(* IEC 61131-3 sources: Elmo_Master/Lasal_PRG/Elmo_EtherCAT_Test_4Axis/Class/_TCPIPServer, 1 file *)

(* ---- _TCPIPServer.st ---- *)
  #ifndef OS_VERSION_MIN_SALAMANDER
    #define OS_VERSION_MIN_SALAMANDER          0x9000
  #endif
  #define TCP_SVR_NO_ERROR                          0

  #define TCP_SVR_ERR_INVALID_SOCKET            -1

  #define TCP_SVR_ERR_SET_PARA_INVALID_CMD     -10
  #define TCP_SVR_ERR_SET_PARA_INVALID_SUB_CMD -11

  #define TCP_SVR_ERR_TASK_ALREADY_EXIST       -12

  // - RETURN VALUES PRIVATE METHOD Read_AP_TaskPeriod
  #define TCP_SVR_ERR_TASK_TIME_NO_APP            -31
  #define TCP_SVR_ERR_TASK_TIME_WRONG_TASK_TYPE   -33
  #define TCP_SVR_ERR_TASK_TIME_OBJ_NOT_FOUND     -35

  // - RETURN VALUES PRIVATE METHOD Read_LSLOBJ_CRC32
  #define TCP_SVR_ERR_GET_LSLOBJ_NAME             -20
  #define TCP_SVR_ERR_INVALID_POINTER             -21

  // - RETURN VALUES PRIVATE METHOD AP_TaskCreate
  #define TCP_SVR_ERR_TASK_CREATE                 -40

  // - RETURN VALUES PRIVATE METHOD AP_SemaCreate
  #define TCP_SVR_ERR_SEMA_CREATE                 -50
  #define TCP_SVR_ERR_SEMA_INVALID_IDX            -51
  #define TCP_SVR_ERR_SEMA_INVALID_NAME           -52

  #define TCP_SVR_SEND_BUFFER_EMPTY               -6
  #define TCP_SVR_ERR_SEND_BUFFER_FATAL_ERROR     -7

  #define TCP_SVR_SEND_BUFFER_FULL      -4

  #define TCP_SVR_SOCK_INFO_CONNECT                 1
  #define TCP_SVR_SOCK_INFO_DISCONNECT              0

  #define TCP_SVR_ERR_GROUP_OS                      0
  #define TCP_SVR_ERR_GROUP_AP                      1

  #define TCP_SVR_ERR_CODE_AP_TIMEOUT              -1

  #ifndef INIT_FIRSTSCAN
    #define INIT_FIRSTSCAN                         12
  #endif

  #ifndef AP_TASK_PRIORITY_DEFAULT
    #define AP_TASK_PRIORITY_DEFAULT               14
  #endif

  #define TCP_SVR_ERR_MAIN_INIT                   -90

  #define TCP_SVR_ERR_MAX_CONN                    -80

  #ifndef KEEPALIVE_INTERVAL_DEFAULT
    #define KEEPALIVE_INTERVAL_DEFAULT           7200
  #endif

  #ifndef KEEPALIVE_RETRYTIME_DEFAULT
    #define KEEPALIVE_RETRYTIME_DEFAULT            75
  #endif

  #ifndef KEEPALIVE_RETRYCNT_DEFUALT
    #define KEEPALIVE_RETRYCNT_DEFUALT             10
  #endif

  #ifndef CLOSE_SOCKET_TYPE_DEFAULT
    #define CLOSE_SOCKET_TYPE_DEFAULT               0
  #endif

#include "..\..\Class\_TCPIPServer\_TCPIPServer.h"
#include "..\..\Class\_TCPIPServer\SalamanderDelay.h"

(*!
<Class
	Name               = "_TCPIPServer"
	Revision           = "1.2"
	RealtimeTask       = "false"
	CyclicTask         = "true"
	DefCyclictime      = "10 ms"
	BackgroundTask     = "false"
	DefBackground      = "always"
	Sigmatek           = "true"
	OSInterface        = "false"
	HighPriority       = "false"
	Automatic          = "false"
	UpdateMode         = "Prescan"
	SharedCommandTable = "true"
	Objectsize         = "(590,120)"
	Comment            = "TCP/IP Server for TCP/IP Communication">
	<Channels>
		<Server Name="Control" Visualized="false" Initialize="false" WriteProtected="true" Retentive="false" Comment="shows the actual TCP/IP state"/>
		<Server Name="ErrorCode" Visualized="false" Initialize="false" WriteProtected="true" Retentive="false" Comment="Shows error codes&#13;&#10; 0 ... no error&#13;&#10;-1 ... general error&#13;&#10;-2 ... timeout error&#13;&#10;-3 ... connection closed by client&#13;&#10;-4 ... File open failed&#13;&#10;-5 ... Copy Data from File failed&#13;&#10;-6 ... Sending Data failed&#13;&#10;-7 ... read SendBuffer failed&#13;&#10;-8 ... BackUp- or Restore-Object failed&#13;&#10;-9 ... Pointer to SendBuffer = NIL&#13;&#10;-10... Pointer to Receive Buffer = NIL&#13;&#10;-11... Write into SendBuffer failed&#13;&#10;-12... Set Socket Option failed&#13;&#10;-13... Data is to big to send&#13;&#10;-14... Received Data is too short&#13;&#10;-15... Received Datasize not equal with specified Datasize&#13;&#10;-16... Received Datasize not equal with specified Datasize (too long)&#13;&#10;-99... Allocate Memory failed&#13;&#10;-100 . Search for Semikolon or Carriage Return failed"/>
		<Server Name="SemaName01" Visualized="true" Initialize="false" WriteProtected="true" Retentive="false" Comment="name of mutex to save the internal connection buffer&#13;&#10;&#13;&#10;This name is also listed in PLCTraceView"/>
		<Server Name="SemaName02" Visualized="true" Initialize="false" WriteProtected="true" Retentive="false" Comment="name of mutex to save the internal connection settings (socket options)&#13;&#10;&#13;&#10;This name is also listed in PLCTraceView"/>
		<Server Name="TaskName" Visualized="true" Initialize="false" WriteProtected="true" Retentive="false" Comment="shows task information&#13;&#10;-) use object in cyclic task&#13;&#10;-) use object in async task&#13;&#10;-) task deactivated&#13;&#10;-) async task error status (error creating async task)&#13;&#10;&#13;&#10;In case of using the object in async task, this name is also listed in PLCTraceView"/>
		<Client Name="_MultiTask" Required="false" Internal="false" Comment="object channel to OS interface class _MultiTask"/>
		<Client Name="_StdLib" Required="false" Internal="false" Comment="object channel to OS interface class _StdLib"/>
		<Client Name="_TaskObjectControl" Required="false" Internal="false" Comment="object channel to OS interface class _TaskObjectControl"/>
		<Client Name="CheckSum" Required="true" Internal="true"/>
		<Client Name="Config" Required="false" Internal="false" Comment="object configuration&#13;&#10;bit0 ... task configuration&#13;&#10;0 = use object in cyclic task&#13;&#10;1 = use object in async task"/>
		<Client Name="ConnectionsPerRun" Required="true" Internal="false" DefValue="1" Comment="Number of connections to process every cycle:&#13;&#10;&#13;&#10;0, 1 = 1 connection per cycle&#13;&#10;2 = 2 connections per cycle&#13;&#10;... up to ...&#13;&#10;&quot;MaxConnections&quot; = all connections every cycle"/>
		<Client Name="MaxConnections" Required="true" Internal="false" DefValue="0" Comment="Maximal number of connections. Maximal possible connections are 128.&#13;&#10;&#13;&#10;0 = 16 connections, because of compatibility to older versions."/>
		<Client Name="Port" Required="true" Internal="false" Comment="port number&#13;&#10;"/>
		<Client Name="SigCLib" Required="false" Internal="false" Comment="object channel to OS interface class SigCLib"/>
		<Client Name="SizeOfTXBuffer" Required="false" Internal="false" Comment="size of TX buffer [byte]&#13;&#10;if 0 there will be 1024 Byte allocated"/>
		<Client Name="StrSemaName01" Required="true" Internal="true"/>
		<Client Name="StrSemaName02" Required="true" Internal="true"/>
		<Client Name="StrTaskName" Required="true" Internal="true"/>
		<Client Name="Timeout" Required="false" Internal="false" Comment="TCP timeout [ms]&#13;&#10;if 0 then Timeout is deactivated"/>
	</Channels>
	<Dependencies>
		<Files>
			<File Path=".\lsl_st_tcp_user.h" Include="false"/>
			<File Path=".\Class\_TCPIPServer\_TCPIPServer.h" Include="true"/>
			<File Path=".\Class\_TCPIPServer\SalamanderDelay.h" Include="true"/>
		</Files>
	</Dependencies>
	<RevDoku>
		<Owner Company="SIGMATEK"/>
		<Dokumentation Revision="1.2" Date="2024-07-01" Author="zoepat" Company="Sigmatek" Description="- increased maximum connections from 16 to 128.&#13;&#10;- added configuration to define the number of connections to be processed per cycle."/>
		<Dokumentation Revision="1.1" Date="2023-03-23" Author="obechr" Company="Sigmatek" Description="changed comments of parameters for method SendData()"/>
		<Dokumentation Revision="1.0" Date="2019-01-15" Author="hoeant" Company="Sigmatek" Description="creation of class"/>
	</RevDoku>
	<Network Name="_TCPIPServer">
		<!-- List of Components in this network -->
		<Components>
			<Object
				Name       = "CheckSum"
				Class      = "_CheckSum"
				Position   = "(240,180)"
				Visualized = "false">
				<Channels>
					<Server Name="ClassSvr"/>
				</Channels>
			</Object>
			<Object
				Name       = "StrSemaName01"
				Class      = "String"
				Position   = "(240,510)"
				Visualized = "true"
				Remotely   = "true">
				<Channels>
					<Server Name="Data"/>
					<Client Name="SingleRealloc" Value="1"/>
				</Channels>
			</Object>
			<Object
				Name       = "StrSemaName02"
				Class      = "String"
				Position   = "(240,660)"
				Visualized = "true"
				Remotely   = "true">
				<Channels>
					<Server Name="Data"/>
					<Client Name="SingleRealloc" Value="1"/>
				</Channels>
			</Object>
			<Object
				Name       = "StrTaskName"
				Class      = "String"
				Position   = "(240,360)"
				Visualized = "true"
				Remotely   = "true">
				<Channels>
					<Server Name="Data"/>
					<Client Name="SingleRealloc" Value="1"/>
				</Channels>
			</Object>
		</Components>
		<Comments>
		</Comments>
		<!-- List of Connections in this network -->
		<Connections>
			<Connection Source="this.CheckSum" Destination="CheckSum.ClassSvr"/>
			<Connection Source="this.StrTaskName" Destination="StrTaskName.Data"/>
			<Connection Source="this.StrSemaName01" Destination="StrSemaName01.Data"/>
			<Connection Source="this.StrSemaName02" Destination="StrSemaName02.Data"/>
			<Connection Source="this.TaskName" Destination="StrTaskName.Data" Vertices="(1028,330),(556,450),"/>
			<Connection Source="this.SemaName01" Destination="StrSemaName01.Data" Vertices="(1028,390),(556,600),"/>
			<Connection Source="this.SemaName02" Destination="StrSemaName02.Data" Vertices="(1028,450),(556,750),"/>
		</Connections>
		<!-- Headerfiles -->
		<Options>
		</Options>
	</Network>
</Class>
*)
_TCPIPServer : CLASS
	TYPE
#pragma pack(push, 1)
	  _BUFFER : STRUCT  //! <Type Comment="Struct for Receive- and Send-Buffer" Name="_BUFFER"/>
	    udSize : UDINT;  //! <Type Comment="Size of Data" Name="_BUFFER.udSize"/>
	    pData : ^void;  //! <Type Comment="Pointer to Data" Name="_BUFFER.pData"/>
	  END_STRUCT;
#pragma pack(pop)
#pragma pack(push, 1)
	  _BUFFER_HEADER : STRUCT
	    DataSize : UDINT;
	  END_STRUCT;
#pragma pack(pop)
	  _FSM_TCPIP_SERVER :  //! <Type Public="true" Comment="stepping switch for TCP/IP connection" Name="_FSM_TCPIP_SERVER"/>
	  (
	    _STATE_NONE,
	    _STATE_INIT_SERVER,
	    _STATE_NO_USER_INTERFACE_CONNECTED,
	    _STATE_IDLE,
	    _STATE_MAIN_SOCK,
	    _STATE_LISTEN,
	    _STATE_ACCEPT,
	    _STATE_CONNECT,
	    _STATE_RECV,
	    _STATE_SHUTDOWN,
	    _STATE_CLOSE_MAIN_SOCK,
	    _STATE_CLOSE_SOCK,
	    _STATE_ERROR,
	    _STATE_ERROR_ALLOCATING_MEMORY,
	    _STATE_ERROR_CREATING_MUTEX,
	    _STATE_ERROR_CREATING_TASK,
	    _STATE_SEND,
	    _STATE_MAIN_SOCK_OPT,
	    _STATE_DEL_CONNECTION,
	    _STATE_CONN_SOCK_OPT
	  )$UDINT;
#pragma pack(push, 1)
	  _TX_RINGBUFFER : STRUCT  //! <Type Comment="struct to handle a ringbuffer" Name="_TX_RINGBUFFER"/>
	    udSize : UDINT;
	    udUsed : UDINT;
	    pMem : ^void;
	    pRead : ^CHAR;
	    pWrite : ^CHAR;
	  END_STRUCT;
#pragma pack(pop)
	  _SocketOptions : BDINT
	  [
	    1 Nagle,
	    2 KeepAlive,
	    3 DelayedAck,
	    4 ReuseAddr,
	    5 Bit5,
	    6 Bit6,
	    7 Bit7,
	    8 Bit8,
	    9 Bit9,
	    10 Bit10,
	    11 Bit11,
	    12 Bit12,
	    13 Bit13,
	    14 Bit14,
	    15 Bit15,
	    16 Bit16,
	    17 Bit17,
	    18 Bit18,
	    19 Bit19,
	    20 Bit20,
	    21 Bit21,
	    22 Bit22,
	    23 Bit23,
	    24 Bit24,
	    25 Bit25,
	    26 Bit26,
	    27 Bit27,
	    28 Bit28,
	    29 Bit29,
	    30 Bit30,
	    31 Bit31,
	    32 Bit32,
	  ];
#pragma pack(push, 1)
	  _KeepAlivePara : STRUCT
	    keepIDLE : DINT;
	    keepINTVL : DINT;
	    keepCNT : DINT;
	  END_STRUCT;
#pragma pack(pop)
#pragma pack(push, 1)
	  _CONNECTION : STRUCT
	    dSocket : DINT;
	    FSM_TCP : _FSM_TCPIP_SERVER;
	    udTimeStamp : UDINT;
	    SendBuffer : _TX_RINGBUFFER;
	    pBufferWaitForSendig : ^CHAR;
	    pBufferWaitForSendingHelp : ^CHAR;
	    BufferHeader : _BUFFER_HEADER;
	    ConnSockOpt : _SocketOptions;
	    pNextConn : ^_CONNECTION;
	    bdSettings : BDINT
	    [
	      1 SockOptChanged,
	      2 Bit2,
	      3 Bit3,
	      4 Bit4,
	      5 Bit5,
	      6 Bit6,
	      7 Bit7,
	      8 Bit8,
	      9 Bit9,
	      10 Bit10,
	      11 Bit11,
	      12 Bit12,
	      13 Bit13,
	      14 Bit14,
	      15 Bit15,
	      16 Bit16,
	      17 Bit17,
	      18 Bit18,
	      19 Bit19,
	      20 Bit20,
	      21 Bit21,
	      22 Bit22,
	      23 Bit23,
	      24 Bit24,
	      25 Bit25,
	      26 Bit26,
	      27 Bit27,
	      28 Bit28,
	      29 Bit29,
	      30 Bit30,
	      31 Bit31,
	      32 Bit32,
	    ];
	    KeepAlivePara : _KeepAlivePara;
	    CloseSocketType : UDINT;
	  END_STRUCT;
#pragma pack(pop)
#pragma pack(push, 1)
	  _KeepAliveParaLasalOS : STRUCT
	    interval : UINT;
	    retry : UINT;
	    timeout : UINT;
	  END_STRUCT;
#pragma pack(pop)
	END_TYPE
  //Servers:
	Control 	: SvrChCmd__FSM_TCPIP_SERVER_PTofCls__TCPIPServer;
	ErrorCode 	: SvrCh_DINT;
	TaskName 	: SvrCh_UDINT;
	SemaName01 	: SvrCh_UDINT;
	SemaName02 	: SvrCh_UDINT;
  //Clients:
	Port 	: CltCh_DINT;
	Timeout 	: CltCh_DINT;
	SizeOfTXBuffer 	: CltCh_UDINT;
	MaxConnections 	: CltCh_DINT;
	ConnectionsPerRun 	: CltCh_DINT;
	Config 	: CltCh_DINT;
	_StdLib 	: CltChCmd__StdLib;
	_MultiTask 	: CltChCmd__MultiTask;
	SigCLib 	: CltChCmd_SigCLib;
	CheckSum 	: CltChCmd__CheckSum;
	StrTaskName 	: CltChCmd_String;
	StrSemaName01 	: CltChCmd_String;
	StrSemaName02 	: CltChCmd_String;
	_TaskObjectControl 	: CltChCmd__TaskObjectControl;
  //Variables:
		dMainSock 	: DINT;			//! <Variable Comment="main socket for TCP/IP connection" Name="dMainSock"/>
		FSM_TCP 	: _FSM_TCPIP_SERVER;			//! <Variable Comment="finite state machine for TCP/IP connection" Name="FSM_TCP"/>
		SocketArray : ARRAY [0..127] OF _CONNECTION;
			//! <Variable Comment="Saves the Informations for each Connection" Name="SocketArray"/>
		RECVbuffer 	: _BUFFER;			//! <Variable Comment="struct of Receive buffer" Name="RECVbuffer"/>
		lsl_tcp_user 	: ^LSL_TCP_USER;
		usInit 	: USINT;
		bdStatus : BDINT
		[
		  1 SalamanderOS,
		  5 CIL_tcp_user,
		  6 CIL_ssl_user,
		  7 CIL_debug,
		  9 InhibNextConn,
		  13 LSLOBJ_CRC32,
		  14 AP_TaskPeriod,
		  15 CyclicTask,
		  16 AsyncTask,
		  17 Sema01,
		  18 Sema02,
		  25 ErrAsyncTask,
		  26 ErrSema01,
		  27 ErrSema02,
		  28 ErrMem,
		  29 ErrorNoUserInterface,
		];

		MaxConn 	: DINT;
		lsl_ssl_user 	: ^LSL_SSL_USER;
		pCIL_DEBUG 	: ^OS_SALAMANDERDEBUG;
		MainSockOpt 	: _SocketOptions;
		AP_TaskTime 	: UDINT;
		AP_TaskHandle 	: MT_TASKHANDLE;
		AP_SemaHandle1 	: MT_SEMAHANDLE;
		AP_SemaSockOpt 	: MT_SEMAHANDLE;
		ActConn 	: DINT;
		pActConn 	: ^_CONNECTION;
		udTimeStamp 	: UDINT;
		udTimeAccept 	: UDINT;
		AP_TaskPriority 	: UDINT;
		KeepAlivePara 	: _KeepAlivePara;
		CloseSocketType 	: UDINT;
		dNewSock 	: DINT;
		pThisInterface 	: ^_TCPIPServerInterface;
  //Functions:
				//! <Function Comment="-) initialize TCP USER pointer to use OS TCP FUNCTIONS&#13;&#10;-) read port number&#13;&#10;-) Allocate Memory for Buffers" Name="Init"/>
	FUNCTION VIRTUAL GLOBAL Init;
				//! <Function Comment="cyclic tast methode which is called if client &#13;&#10;cConfig = 0" Name="CyWork"/>
	FUNCTION VIRTUAL GLOBAL CyWork
		VAR_INPUT
			EAX 	: UDINT;
		END_VAR
		VAR_OUTPUT
			state (EAX) 	: UDINT;
		END_VAR;
				//! <Function Comment="this function writes data into the TX buffer&#13;&#10;" Name="SENDbuffer_Write"/>
	FUNCTION SENDbuffer_Write
		VAR_INPUT
			pData 	: ^void;
			udSize 	: UDINT;
			pBuffer 	: ^_TX_RINGBUFFER;
		END_VAR
		VAR_OUTPUT
			dRetcode 	: DINT;
		END_VAR;
				//! <Function Comment="Function to send data over TCP/IP&#13;&#10;&#13;&#10;--------------------------------------&#13;&#10;Input variables&#13;&#10;--------------------------------------&#13;&#10;-) pData ... pointer to data to send&#13;&#10;-) udSize ... size of data to send [byte]&#13;&#10;-) dSock ... Receiver-Socket&#13;&#10;&#13;&#10;--------------------------------------&#13;&#10;Output variables&#13;&#10;--------------------------------------&#13;&#10;-) dRetcode&#13;&#10;   &lt; 0:&#13;&#10;      -1 ... TCP Client not ready&#13;&#10;      else ... OS TCP error code&#13;&#10;&#13;&#10;   &gt;=0:&#13;&#10;      dRetcode = udSize ... Sending data over TCP/IP successful" Name="SendTCP"/>
	FUNCTION SendTCP
		VAR_INPUT
			pData 	: ^void;
			udSize 	: UDINT;
			dSock 	: DINT;
			bDirect 	: DINT;
		END_VAR
		VAR_OUTPUT
			dRetcode 	: DINT;
		END_VAR;
				//! <Function Comment="Handles the Connection and Data receiving and sending" Name="CyclicCall"/>
	FUNCTION VIRTUAL GLOBAL CyclicCall;
				//! <Function Comment="Read Send Buffer" Name="SENDbuffer_Read"/>
	FUNCTION SENDbuffer_Read
		VAR_INPUT
			pBuffer 	: ^_TX_RINGBUFFER;
			pData 	: ^void;
			udSize 	: UDINT;
		END_VAR
		VAR_OUTPUT
			Retcode 	: DINT;
		END_VAR;
				//! <Function Comment="Send Data over TCP/IP" Name="SendData"/>
	FUNCTION VIRTUAL GLOBAL SendData
		VAR_INPUT
			pData 	: ^void;			//! <Variable Comment="Pointer to Data" Name="SendData.pData"/>
			udSize 	: UDINT;			//! <Variable Comment="Size of Data" Name="SendData.udSize"/>
			dSock 	: DINT;			//! <Variable Comment="Socket to which it should be send" Name="SendData.dSock"/>
			bDirect 	: BOOL;			//! <Variable Comment="0 ... Write it to Send Buffer and send it in next Cyclus&#13;&#10;1 ... Send it imediatly" Name="SendData.bDirect"/>
		END_VAR
		VAR_OUTPUT
			dRetcode 	: DINT;			//! <Variable Comment="&gt;=0 .. size of the processed data&#13;&#10;&lt;0 ..  error occured" Name="SendData.dRetcode"/>
		END_VAR;

	FUNCTION Read_LSLOBJ_CRC32
		VAR_INPUT
			pCRC32 	: ^CHAR;
		END_VAR
		VAR_OUTPUT
			Retcode 	: DINT;
		END_VAR;

	FUNCTION Read_AP_TaskPeriod
		VAR_OUTPUT
			Retcode 	: DINT;
		END_VAR;

	FUNCTION AP_TaskCreate
		VAR_INPUT
			pTaskName 	: ^CHAR;
			pCallback 	: ^void;
		END_VAR
		VAR_OUTPUT
			Retcode 	: DINT;
		END_VAR;

	FUNCTION AP_TaskCallback
		VAR_INPUT
			Param0 	: ^void;
		END_VAR;

	FUNCTION GetMultiTaskErrorCode
		VAR_INPUT
			pErrTxt 	: ^CHAR;
		END_VAR;

	FUNCTION AP_SemaCreate
		VAR_INPUT
			pSemaName 	: ^CHAR;
			Index 	: DINT;
		END_VAR
		VAR_OUTPUT
			Retcode 	: DINT;
		END_VAR;

	FUNCTION AP_TaskDelay
		VAR_INPUT
			udTaskDelay 	: UDINT;
		END_VAR;

	FUNCTION SetMainSocketOptions
		VAR_OUTPUT
			Retcode 	: DINT;
		END_VAR;

	FUNCTION RingbufferReadEntry
		VAR_INPUT
			pBuffer 	: ^_TX_RINGBUFFER;
			pData 	: ^void;
			pSize 	: ^UDINT;
		END_VAR
		VAR_OUTPUT
			Retcode 	: DINT;
		END_VAR;

	FUNCTION RingbufferWriteEntry
		VAR_INPUT
			pBuffer 	: ^_TX_RINGBUFFER;
			pData 	: ^void;
			udSize 	: UDINT;
		END_VAR
		VAR_OUTPUT
			Retcode 	: DINT;
		END_VAR;

	FUNCTION AP_SemaWait
		VAR_INPUT
			SemaHandle 	: MT_SEMAHANDLE;
		END_VAR;

	FUNCTION AP_SemaSignal
		VAR_INPUT
			SemaHandle 	: MT_SEMAHANDLE;
		END_VAR;

	FUNCTION SetSocketOptions
		VAR_INPUT
			pConn 	: ^_CONNECTION;
		END_VAR
		VAR_OUTPUT
			Retcode 	: DINT;
		END_VAR;

	FUNCTION AddConnIntern
		VAR_INPUT
			dSocket 	: DINT;
			ppConn 	: ^pVoid;
		END_VAR
		VAR_OUTPUT
			Retcode 	: DINT;
		END_VAR;

	FUNCTION DelConnIntern
		VAR_INPUT
			dSocket 	: DINT;
		END_VAR
		VAR_OUTPUT
			Retcode 	: DINT;
		END_VAR;
				//! <Function Comment="method is called with socket informations of the connection sockets" Name="ConnSocketInfo"/>
	FUNCTION ConnSocketInfo
		VAR_INPUT
			dSock 	: DINT;			//! <Variable Comment="socket number" Name="ConnSocketInfo.dSock"/>
			InfoPara1 	: DINT;			//! <Variable Comment="0 ... socket disconnected&#13;&#10;1 ... socket connected" Name="ConnSocketInfo.InfoPara1"/>
			InfoPara2 	: DINT;			//! <Variable Comment="InfoPara2 = 0" Name="ConnSocketInfo.InfoPara2"/>
		END_VAR;
				//! <Function Comment="method is called with socket error status of the connection sockets&#13;&#10;&#13;&#10;-) TCP error (callback: ErrorGroup = 0, ErrorCode = TCP error status)&#13;&#10;-) error code definition in lsl_st_tcp_user.h&#13;&#10;&#13;&#10;-)  internal error (callback: ErrorGroup = 1, ErrorCode = internal error status)&#13;&#10;-) -1: receive timeout (in case of timeout is set)" Name="ConnSocketError"/>
	FUNCTION ConnSocketError
		VAR_INPUT
			dSock 	: DINT;			//! <Variable Comment="socket number" Name="ConnSocketError.dSock"/>
			FSM_TCP 	: _FSM_TCPIP_SERVER;			//! <Variable Comment="status of the state machine of the connection socket" Name="ConnSocketError.FSM_TCP"/>
			ErrGroup 	: DINT;			//! <Variable Comment="0 ... OS error (OS_TCP_USER)&#13;&#10;1 ... AP error (connection timeout)" Name="ConnSocketError.ErrGroup"/>
			ErrCode 	: DINT;			//! <Variable Comment="ErrGroup = 0 (OS error)&#13;&#10;ErrCode definition in lsl_st_tcp_user.h&#13;&#10;&#13;&#10;ErrGroup = 1 (AP error)&#13;&#10;ErrCode = -1 ... connection timeout&#13;&#10;" Name="ConnSocketError.ErrCode"/>
		END_VAR;
				//! <Function Comment="method is called with socket informations of the main socket" Name="MainSocketError"/>
	FUNCTION MainSocketError
		VAR_INPUT
			FSM_TCP 	: _FSM_TCPIP_SERVER;			//! <Variable Comment="status of the state machine of the main socket" Name="MainSocketError.FSM_TCP"/>
			ErrGroup 	: DINT;			//! <Variable Comment="0 ... OS error (OS_TCP_USER)" Name="MainSocketError.ErrGroup"/>
			ErrCode 	: DINT;
		END_VAR;
				//! <Function Comment="Method to set main parameters. Main parameters will be used for every new connection." Name="SetMainParameter"/>
	FUNCTION VIRTUAL GLOBAL SetMainParameter
		VAR_INPUT
			Cmd 	: DINT;			//! <Variable Comment="0 ... (SVR_TCP_CMD_SETSOCKOPT) socket option&#13;&#10;1 ... (SVR_TCP_CMD_TASKPRIO) task priority of async task (in case of using object in async task)&#13;&#10;2 ... (SVR_TCP_CMD_CLOSESOCKETTYPE) close socket type&#13;&#10;3 ... (SVR_TCP_CMD_KEEPALIVEPARA) keep alive parameter&#13;&#10;" Name="SetMainParameter.Cmd"/>
			SubCmd 	: DINT;			//! <Variable Comment="Cmd = 0 (SVR_TCP_CMD_SETSOCKOPT)&#13;&#10;-) SubCmd = 0:  SVR_TCP_SOCKOPT_NAGLE ... activate/deactivate nagle algorithm&#13;&#10;-) SubCmd = 1:  SVR_TCP_SOCKOPT_KEEPALIVE ... activate/deactivate keepalive message&#13;&#10;-) SubCmd = 2:  SVR_TCP_SOCKOPT_DELAYEDACK ... activate/deactivate delayed acknowledge packet&#13;&#10;-) SubCmd = 3:  SVR_TCP_SOCKOPT_REUSEADDR ... activate/deactivate option reuse address&#13;&#10;&#13;&#10;Cmd = 1 (SVR_TCP_CMD_TASKPRIO)&#13;&#10;-) SubCmd = 0: task priority of async task&#13;&#10;&#13;&#10;&#13;&#10;Cmd = 2 (SVR_TCP_CMD_CLOSESOCKETTYPE)&#13;&#10;-) SubCmd = 0: SVR_TCP_CLOSESOCKETTYPE&#13;&#10;&#13;&#10;Cmd = 3 (SVR_TCP_CMD_KEEPALIVEPARA)&#13;&#10;-) SubCmd = 0:  SVR_TCP_KEEPALIVE_KEEPIDLE&#13;&#10;-) SubCmd = 1:  SVR_TCP_KEEPALIVE_KEEPINTVL&#13;&#10;-) SubCmd = 2:  SVR_TCP_KEEPALIVE_KEEPCNT&#13;&#10;" Name="SetMainParameter.SubCmd"/>
			ParaValue 	: DINT;			//! <Variable Comment="Cmd = 0 (SVR_TCP_CMD_SETSOCKOPT)&#13;&#10;-) 1 ... Activate option&#13;&#10;-) 0 ... Deactivate option&#13;&#10;&#13;&#10;Cmd = 1 (SVR_TCP_CMD_TASKPRIO)&#13;&#10;-) task priority 1-14&#13;&#10;&#13;&#10;Cmd = 2 (SVR_TCP_CMD_CLOSESOCKETTYPE)&#13;&#10;-) 0 ... Graceful Close&#13;&#10;-) 1 ... Hard Close&#13;&#10;&#13;&#10;Cmd = 3 (SVR_TCP_CMD_KEEPALIVEPARA)&#13;&#10;-)SubCmd = 0: Interval time [ms] for the Keep Alive packages&#13;&#10;-)SubCmd = 1: Retry time [ms] of Keep Alive packages&#13;&#10;-)SubCmd = 2: Define how often the retry will be attempted. Retry time * Retry Count = timeout for Keep Alive packages" Name="SetMainParameter.ParaValue"/>
		END_VAR
		VAR_OUTPUT
			Retcode 	: DINT;			//! <Variable Comment="0 ... success&#13;&#10;-10 ... invalid CMD&#13;&#10;-11 ... invalid SubCMD&#13;&#10;-12 ... error set task priority - task already created&#13;&#10;-90 ... object not initialized (initialization in first Init() call)" Name="SetMainParameter.Retcode"/>
		END_VAR;
				//! <Function Comment="method to read main parameters" Name="ReadMainParameter"/>
	FUNCTION VIRTUAL GLOBAL ReadMainParameter
		VAR_INPUT
			Cmd 	: DINT;			//! <Variable Comment="0 ... (SVR_TCP_CMD_SETSOCKOPT) socket option&#13;&#10;1 ... (SVR_TCP_CMD_TASKPRIO) task priority of async task (in case of using object in async task)&#13;&#10;2 ... (SVR_TCP_CMD_CLOSESOCKETTYPE) close socket type&#13;&#10;3 ... (SVR_TCP_CMD_KEEPALIVEPARA) keep alive parameter" Name="ReadMainParameter.Cmd"/>
			SubCmd 	: DINT;			//! <Variable Comment="Cmd = 0 (SVR_TCP_CMD_SETSOCKOPT)&#13;&#10;-) SubCmd = 0:  SVR_TCP_SOCKOPT_NAGLE ... activate/deactivate nagle algorithm&#13;&#10;-) SubCmd = 1:  SVR_TCP_SOCKOPT_KEEPALIVE ... activate/deactivate keepalive message&#13;&#10;-) SubCmd = 2:  SVR_TCP_SOCKOPT_DELAYEDACK ... activate/deactivate delayed acknowledge packet&#13;&#10;-) SubCmd = 3:  SVR_TCP_SOCKOPT_REUSEADDR ... activate/deactivate option reuse address&#13;&#10;&#13;&#10;Cmd = 1 (SVR_TCP_CMD_TASKPRIO)&#13;&#10;-) SubCmd = 0: task priority of async task&#13;&#10;&#13;&#10;&#13;&#10;Cmd = 2 (SVR_TCP_CMD_CLOSESOCKETTYPE)&#13;&#10;-) SubCmd = 0: SVR_TCP_CLOSESOCKETTYPE&#13;&#10;&#13;&#10;Cmd = 3 (SVR_TCP_CMD_KEEPALIVEPARA)&#13;&#10;-) SubCmd = 0:  SVR_TCP_KEEPALIVE_KEEPIDLE&#13;&#10;-) SubCmd = 1:  SVR_TCP_KEEPALIVE_KEEPINTVL&#13;&#10;-) SubCmd = 2:  SVR_TCP_KEEPALIVE_KEEPCNT&#13;&#10;" Name="ReadMainParameter.SubCmd"/>
			pParaValue 	: ^DINT;			//! <Variable Comment="pointer to target parameter value" Name="ReadMainParameter.pParaValue"/>
		END_VAR
		VAR_OUTPUT
			Retcode 	: DINT;			//! <Variable Comment="0 ... success&#13;&#10;-10 ... invalid CMD&#13;&#10;-11 ... invalid SubCMD&#13;&#10;-90 ... object not initialized (initialization in first Init() call)" Name="ReadMainParameter.Retcode"/>
		END_VAR;
				//! <Function Comment="method to set connection socket parameters" Name="SetSocketParameter"/>
	FUNCTION VIRTUAL GLOBAL SetSocketParameter
		VAR_INPUT
			dSock 	: DINT;			//! <Variable Comment="socket number" Name="SetSocketParameter.dSock"/>
			Cmd 	: DINT;			//! <Variable Comment="0 ... (SVR_TCP_CMD_SETSOCKOPT) socket option&#13;&#10;2 ... (SVR_TCP_CMD_CLOSESOCKETTYPE) close socket type&#13;&#10;3 ... (SVR_TCP_CMD_KEEPALIVEPARA) keep alive parameter" Name="SetSocketParameter.Cmd"/>
			SubCmd 	: DINT;			//! <Variable Comment="Cmd = 0 (SVR_TCP_CMD_SETSOCKOPT)&#13;&#10;-) SubCmd = 0:  SVR_TCP_SOCKOPT_NAGLE ... activate/deactivate nagle algorithm&#13;&#10;-) SubCmd = 1:  SVR_TCP_SOCKOPT_KEEPALIVE ... activate/deactivate keepalive message&#13;&#10;-) SubCmd = 2:  SVR_TCP_SOCKOPT_DELAYEDACK ... activate/deactivate delayed acknowledge packet&#13;&#10;-) SubCmd = 3:  SVR_TCP_SOCKOPT_REUSEADDR ... activate/deactivate option reuse address&#13;&#10;&#13;&#10;Cmd = 2 (SVR_TCP_CMD_CLOSESOCKETTYPE)&#13;&#10;-) SubCmd = 0: SVR_TCP_CLOSESOCKETTYPE&#13;&#10;&#13;&#10;Cmd = 3 (SVR_TCP_CMD_KEEPALIVEPARA)&#13;&#10;-) SubCmd = 0:  SVR_TCP_KEEPALIVE_KEEPIDLE&#13;&#10;-) SubCmd = 1:  SVR_TCP_KEEPALIVE_KEEPINTVL&#13;&#10;-) SubCmd = 2:  SVR_TCP_KEEPALIVE_KEEPCNT&#13;&#10;" Name="SetSocketParameter.SubCmd"/>
			ParaValue 	: DINT;			//! <Variable Comment="Cmd = 0 (socket option)&#13;&#10;-) 1 ... Activate option&#13;&#10;-) 0 ... Deactivate option&#13;&#10;&#13;&#10;Cmd = 2 (SVR_TCP_CMD_CLOSESOCKETTYPE)&#13;&#10;-) 0 ... Graceful Close&#13;&#10;-) 1 ... Hard Close&#13;&#10;&#13;&#10;Cmd = 3 (SVR_TCP_CMD_KEEPALIVEPARA)&#13;&#10;-)SubCmd = 0: Interval time [ms] for the Keep Alive packages&#13;&#10;-)SubCmd = 1: Retry time [ms] of Keep Alive packages&#13;&#10;-)SubCmd = 2: Define how often the retry will be attempted. Retry time * Retry Count = timeout for Keep Alive packages" Name="SetSocketParameter.ParaValue"/>
		END_VAR
		VAR_OUTPUT
			Retcode 	: DINT;			//! <Variable Comment="0 ... success&#13;&#10;-1 ... invalid socket number&#13;&#10;-10 ... invalid CMD&#13;&#10;-11 ... invalid SubCMD" Name="SetSocketParameter.Retcode"/>
		END_VAR;
				//! <Function Comment="method to read connection socket parameters" Name="ReadSocketParameter"/>
	FUNCTION VIRTUAL GLOBAL ReadSocketParameter
		VAR_INPUT
			dSock 	: DINT;			//! <Variable Comment="socket number" Name="ReadSocketParameter.dSock"/>
			Cmd 	: DINT;			//! <Variable Comment="0 ... (SVR_TCP_CMD_SETSOCKOPT) socket option&#13;&#10;2 ... (SVR_TCP_CMD_CLOSESOCKETTYPE) close socket type&#13;&#10;3 ... (SVR_TCP_CMD_KEEPALIVEPARA) keep alive parameter" Name="ReadSocketParameter.Cmd"/>
			SubCmd 	: DINT;			//! <Variable Comment="Cmd = 0 (SVR_TCP_CMD_SETSOCKOPT)&#13;&#10;-) SubCmd = 0:  SVR_TCP_SOCKOPT_NAGLE ... activate/deactivate nagle algorithm&#13;&#10;-) SubCmd = 1:  SVR_TCP_SOCKOPT_KEEPALIVE ... activate/deactivate keepalive message&#13;&#10;-) SubCmd = 2:  SVR_TCP_SOCKOPT_DELAYEDACK ... activate/deactivate delayed acknowledge packet&#13;&#10;-) SubCmd = 3:  SVR_TCP_SOCKOPT_REUSEADDR ... activate/deactivate option reuse address&#13;&#10;&#13;&#10;Cmd = 2 (SVR_TCP_CMD_CLOSESOCKETTYPE)&#13;&#10;-) SubCmd = 0: SVR_TCP_CLOSESOCKETTYPE&#13;&#10;&#13;&#10;Cmd = 3 (SVR_TCP_CMD_KEEPALIVEPARA)&#13;&#10;-) SubCmd = 0:  SVR_TCP_KEEPALIVE_KEEPIDLE&#13;&#10;-) SubCmd = 1:  SVR_TCP_KEEPALIVE_KEEPINTVL&#13;&#10;-) SubCmd = 2:  SVR_TCP_KEEPALIVE_KEEPCNT&#13;&#10;" Name="ReadSocketParameter.SubCmd"/>
			pParaValue 	: ^DINT;			//! <Variable Comment="pointer to target parameter value" Name="ReadSocketParameter.pParaValue"/>
		END_VAR
		VAR_OUTPUT
			Retcode 	: DINT;			//! <Variable Comment="0 ... success&#13;&#10;-1 ... invalid socket number&#13;&#10;-10 ... invalid CMD&#13;&#10;-11 ... invalid SubCMD" Name="ReadSocketParameter.Retcode"/>
		END_VAR;

	FUNCTION CheckSocketValid
		VAR_INPUT
			dSock 	: DINT;
			ppConn 	: ^pVoid;
		END_VAR
		VAR_OUTPUT
			Retcode 	: BOOL;
		END_VAR;
				//! <Function Comment="Internal Methode to register the Interface Object." Name="AddInterface"/>
	FUNCTION GLOBAL AddInterface
		VAR_INPUT
			thispointer 	: ^void;			//! <Variable Comment="pointer to InterfaceObjekt (this)&#13;&#10;" Name="AddInterface.thispointer"/>
		END_VAR
		VAR_OUTPUT
			dRetcode 	: DINT;			//! <Variable Comment="1..OK (Interface installed )&#13;&#10;-1.. Error (Interface already installed)&#13;&#10;-2.. Error (Pointer not valid)" Name="AddInterface.dRetcode"/>
		END_VAR;
  //Tables:
	FUNCTION @STD
		VAR_OUTPUT
			ret_code	: CONFSTATES;
		END_VAR;
	FUNCTION GLOBAL TAB @CT_;
END_CLASS;

#pragma using _CheckSum
#pragma using String
#pragma usingLtd _MultiTask
#pragma usingLtd _StdLib
#pragma usingLtd _TaskObjectControl
#pragma usingLtd SigCLib

#pragma usingLtd _TCPIPServerInterface

#pragma usingltd _TCPIPServerInterface

FUNCTION VIRTUAL GLOBAL _TCPIPServer::Init
VAR
	i                     : USINT;
  udStrLen              : UDINT;
  dRet                  : DINT;
  szCRC32               : ARRAY [0..15] OF CHAR;
  szTaskName            : ARRAY [0..63] OF CHAR;
  szErrCode             : ARRAY [0..31] OF CHAR;
  szSemaName            : ARRAY [0..63] OF CHAR;
END_VAR

  // -------------------------------------------------------------------------------------------------------
  // -------------------------------------------------------------------------------------------------------
  // - F I R S T   I N I T   R U N   ( M A I N   I N I T )
  // -------------------------------------------------------------------------------------------------------
  // -------------------------------------------------------------------------------------------------------
  FSM_TCP := _STATE_INIT_SERVER;
  if (usInit = 0) then

    // -------------------------------------------------------------------------------------
    // -------------------------------------------------------------------------------------
    // - SET DEFAULT SETTINGS
    // -------------------------------------------------------------------------------------
    // -------------------------------------------------------------------------------------
    MainSockOpt.Nagle      := true;
    MainSockOpt.KeepAlive  := false;
    MainSockOpt.DelayedAck := true;
    MainSockOpt.ReuseAddr  := true;

    AP_TaskPriority         := AP_TASK_PRIORITY_DEFAULT;

    KeepAlivePara.keepIDLE  := KEEPALIVE_INTERVAL_DEFAULT;
    KeepAlivePara.keepINTVL := KEEPALIVE_RETRYTIME_DEFAULT;
    KeepAlivePara.keepCNT   := KEEPALIVE_RETRYCNT_DEFUALT;

    CloseSocketType         := CLOSE_SOCKET_TYPE_DEFAULT;

    // -------------------------------------------------------------------------------------
    // -------------------------------------------------------------------------------------
    // - READ CONFIGURATION PARAMETER
    // -------------------------------------------------------------------------------------
    // -------------------------------------------------------------------------------------
    Port           := Port.Read();
    Config         := Config.Read();
    Timeout        := Timeout.Read();
    MaxConnections := MaxConnections.Read();
    SizeOfTXBuffer := SizeOfTXBuffer.Read();
    ConnectionsPerRun := ConnectionsPerRun.Read();

    // -------------------------------------------------------------------------------------
    // -------------------------------------------------------------------------------------
    // - CHECK GENERAL PARAMETER CONFIGURATION
    // -------------------------------------------------------------------------------------
    // -------------------------------------------------------------------------------------
    if MaxConnections <= 0 then
      MaxConnections := 16;
    elsif MaxConnections > 128 then
      MaxConnections := 128;
    end_if;
    MaxConn := MaxConnections;

    if (SizeOfTXBuffer = 0) then
      SizeOfTXBuffer := 1024;
    end_if;

    //limit between 1 and MaxConnections
    if ConnectionsPerRun <= 0 then
      ConnectionsPerRun := 1;
    elsif ConnectionsPerRun > MaxConnections then
      ConnectionsPerRun := MaxConnections;
    end_if;

    // -------------------------------------------------------------------------------------
    // -------------------------------------------------------------------------------------
    // - READ OS INFORMATION
    // -------------------------------------------------------------------------------------
    // -------------------------------------------------------------------------------------
    if (_RtOSVersion >= OS_VERSION_MIN_SALAMANDER) then
      bdStatus.SalamanderOS := true;
    end_if;

    // -------------------------------------------------------------------------------------
    // -------------------------------------------------------------------------------------
    // - READ OS CIL INTERFACE INFORMATION
    // -------------------------------------------------------------------------------------
    // -------------------------------------------------------------------------------------
    if OS_CILGET("TCP_USER", #lsl_tcp_user) then
      lsl_tcp_user := NIL;
    else
      bdStatus.CIL_tcp_user := true;
    end_if;

    if OS_CILGET("SSL_USER", #lsl_ssl_user) then
      lsl_ssl_user := NIL;
    else
      bdStatus.CIL_ssl_user := true;
    end_if;

    if OS_CILGET("SALAMANDERDEBUG", #pCIL_DEBUG) then
      pCIL_DEBUG := NIL;
    else
      bdStatus.CIL_debug := true;
    end_if;

    // -------------------------------------------------------------------------------------
    // -------------------------------------------------------------------------------------
    // - ALLOCATE MEMORY FOR RECEIVE BUFFER
    // -------------------------------------------------------------------------------------
    // -------------------------------------------------------------------------------------
    RECVbuffer.pData := _StdLib.Malloc(size := to_UDINT(SizeOfTXBuffer));
    if (RECVbuffer.pData = NIL) then
      bdStatus.ErrMem := true;
      ErrorCode := -99;
    end_if;

    // -------------------------------------------------------------------------------------
    // -------------------------------------------------------------------------------------
    // - ALLOCATE MEMORY FOR SEND BUFFER
    // -------------------------------------------------------------------------------------
    // -------------------------------------------------------------------------------------
    for i := 0 to ((MaxConn-1)$USINT) do

      SocketArray[i].dSocket     := 0;
      SocketArray[i].udTimeStamp := 0;
      SocketArray[i].FSM_TCP     := _STATE_IDLE;
      SocketArray[i].pNextConn   := NIL;
      SocketArray[i].SendBuffer.pMem := _StdLib.Malloc(size:=(SizeOfTXBuffer + (10 *sizeof(_BUFFER_HEADER)))); // allocate memory for Ringbuffer (+ 10 * size of Buffer-Header to have enogh Memory)

      if SocketArray[i].SendBuffer.pMem = NIL then
        bdStatus.ErrMem := true;
        ErrorCode := -99;
      else
        SocketArray[i].SendBuffer.pRead  := SocketArray[i].SendBuffer.pMem$^USINT;
        SocketArray[i].SendBuffer.pWrite := SocketArray[i].SendBuffer.pMem$^USINT;
        SocketArray[i].SendBuffer.udSize := SizeOfTXBuffer;
        SocketArray[i].SendBuffer.udUsed := 0;
      end_if;

      SocketArray[i].pBufferWaitForSendig$^void := _StdLib.Malloc(size:=SizeOfTXBuffer); //allocate memory for Sendbuffer

      if SocketArray[i].pBufferWaitForSendig = NIL then
        bdStatus.ErrMem := true;
        ErrorCode := -99;
      end_if;

    end_for;

    // -------------------------------------------------------------------------------------
    // -------------------------------------------------------------------------------------
    // - CHECK USER INTERFACE AVAILABLE
    // -------------------------------------------------------------------------------------
    // -------------------------------------------------------------------------------------

    bdStatus.ErrorNoUserInterface := TRUE;

  end_if;

  usInit += 1;

  // -------------------------------------------------------------------------------------------------------
  // -------------------------------------------------------------------------------------------------------
  // - F I R S T S C A N
  // -------------------------------------------------------------------------------------------------------
  // -------------------------------------------------------------------------------------------------------
  if (_firstscan) then

    // -------------------------------------------------------------------------------------
    // -------------------------------------------------------------------------------------
    // - READ THE LASAL OBJECT CRC32
    // -------------------------------------------------------------------------------------
    // -------------------------------------------------------------------------------------
    dRet := Read_LSLOBJ_CRC32(#szCRC32[0]);
    case dRet of
      (*==================================================================*)
      TCP_SVR_NO_ERROR: // - NO ERROR
      (*==================================================================*)
        bdStatus.LSLOBJ_CRC32 := true;
      (*==================================================================*)
      else // - ERROR WHILE READING THE LASAL OBJECT CRC32 (USE THIS PTR)
      (*==================================================================*)
        SigCLib.IToA(this$DINT, #szCRC32[0], 0x10);
    end_case;

    // -------------------------------------------------------------------------------------
    // -------------------------------------------------------------------------------------
    // - MUTEX CONNECTION INIT
    // -------------------------------------------------------------------------------------
    // -------------------------------------------------------------------------------------
    SigCLib.StrCpy(#szSemaName[0], "USR_SEMA_");
    SigCLib.StrCat(#szSemaName[0], #szCRC32[0]);
    SigCLib.StrCat(#szSemaName[0], "_01");
    dRet := AP_SemaCreate(#szSemaName[4], 0);
    if (dRet = TCP_SVR_NO_ERROR) then
      bdStatus.Sema01 := true;
    else
      bdStatus.ErrSema01 := true;
      GetMultiTaskErrorCode(#szErrCode[0]);
      SigCLib.StrCpy(#szTaskName[0], "SEMA ERR: CREATE SEMA (");
      SigCLib.StrCat(#szTaskName[0], #szErrCode[0]);
      SigCLib.StrCat(#szTaskName[0], ")");
    end_if;

    udStrLen := SigCLib.StrLen(#szSemaName[0]);
    StrSemaName01.WriteDataOff(udStrLen, 0, #szSemaName[0]);

    // -------------------------------------------------------------------------------------
    // -------------------------------------------------------------------------------------
    // - MUTEX SOCKET OPTION INIT
    // -------------------------------------------------------------------------------------
    // -------------------------------------------------------------------------------------
    SigCLib.StrCpy(#szSemaName[0], "USR_SEMA_");
    SigCLib.StrCat(#szSemaName[0], #szCRC32[0]);
    SigCLib.StrCat(#szSemaName[0], "_02");
    dRet := AP_SemaCreate(#szSemaName[4], 1);
    if (dRet = TCP_SVR_NO_ERROR) then
      bdStatus.Sema01 := true;
    else
      bdStatus.ErrSema01 := true;
      GetMultiTaskErrorCode(#szErrCode[0]);
      SigCLib.StrCpy(#szTaskName[0], "SEMA ERR: CREATE SEMA (");
      SigCLib.StrCat(#szTaskName[0], #szErrCode[0]);
      SigCLib.StrCat(#szTaskName[0], ")");
    end_if;

    udStrLen := SigCLib.StrLen(#szSemaName[0]);
    StrSemaName02.WriteDataOff(udStrLen, 0, #szSemaName[0]);

    // -------------------------------------------------------------------------------------
    // -------------------------------------------------------------------------------------
    // - TASK INIT
    // -------------------------------------------------------------------------------------
    // -------------------------------------------------------------------------------------
    udTimeAccept := 500;

    dRet := Read_AP_TaskPeriod();
    if (dRet = TCP_SVR_NO_ERROR) then
      bdStatus.AP_TaskPeriod := true;
      if (Config AND 0x1) then
        // - CYCLIC CALL IN PARALLEL TASK
        SigCLib.StrCpy(#szTaskName[0], "USR_TASK_");
        SigCLib.StrCat(#szTaskName[0], #szCRC32[0]);
        dRet := AP_TaskCreate(#szTaskName[4], #AP_TaskCallback());
        if (dRet = TCP_SVR_NO_ERROR) then
          bdStatus.AsyncTask := true;
        else
          bdStatus.ErrAsyncTask := true;
          GetMultiTaskErrorCode(#szErrCode[0]);
          SigCLib.StrCpy(#szTaskName[0], "TASK ERR: CREATE TASK (");
          SigCLib.StrCat(#szTaskName[0], #szErrCode[0]);
          SigCLib.StrCat(#szTaskName[0], ")");
        end_if;
      else
        // - CYCLIC CALL IN CYCLIC TASK
        bdStatus.CyclicTask := true;
        SigCLib.StrCpy(#szTaskName[0], "CyclicTask");
      end_if;

      // ---------------------------------------------------------------------
      // - ADJUST TIME BETWEEN ACCEPT STEPS FOR COMPATIBILITY
      // ---------------------------------------------------------------------
      if (bdStatus.SalamanderOS = true) then
        udTimeAccept := AP_TaskTime / 1000;
        if (udTimeAccept = 0) then
          udTimeAccept := 1;
        end_if;
      else
        udTimeAccept := AP_TaskTime;
      end_if;
      udTimeAccept := udTimeAccept * 4;

    else

      case dRet of
        (*==================================================================*)
        TCP_SVR_ERR_TASK_TIME_NO_APP:
        (*==================================================================*)
          SigCLib.StrCpy(#szTaskName[0], "TASK ERR: LSLOBJ (NO APPLICATION)");
        (*==================================================================*)
        TCP_SVR_ERR_TASK_TIME_WRONG_TASK_TYPE:
        (*==================================================================*)
          SigCLib.StrCpy(#szTaskName[0], "TASK ERR: LSLOBJ (WRONG TASK TYPE)");
        (*==================================================================*)
        TCP_SVR_ERR_TASK_TIME_OBJ_NOT_FOUND:
        (*==================================================================*)
          SigCLib.StrCpy(#szTaskName[0], "task deactivated");
        (*==================================================================*)
        else
        (*==================================================================*)
          SigCLib.StrCpy(#szTaskName[0], "TASK ERR: LSLOBJ (UNKNOWN ERROR)");
      end_case;

    end_if;

    udStrLen := SigCLib.StrLen(#szTaskName[0]);
    StrTaskName.WriteDataOff(udStrLen, 0, #szTaskName[0]);

  end_if;

END_FUNCTION

FUNCTION VIRTUAL GLOBAL _TCPIPServer::CyWork
	VAR_INPUT
		EAX 	: UDINT;
	END_VAR
	VAR_OUTPUT
		state (EAX) 	: UDINT;
	END_VAR

  if (bdStatus.CyclicTask = true) then
    CyclicCall();
  end_if;

	state := READY;

END_FUNCTION

FUNCTION VIRTUAL GLOBAL _TCPIPServer::CyclicCall
VAR
  dBytes        : DINT;
  i             : DINT;
  dRet          : DINT;
  dAccSock      : DINT;
  pConn         : ^_CONNECTION;
  UserDataToRead : udint;
  ConnPerRun    : DINT;
END_VAR

//++++++++++++++++++++++++++++++++++++++++++++++++++++++++++++++++++++++++++++++++++++++++++++
//++                                                                                        ++
//++    this finite state machine is used for the main TCP/IP connection:                   ++
//++                                                                                        ++
//++    -> allocate sockets                                                                 ++
//++    -> build a connection to a specified socket                                         ++
//++    -> receive data from Client                                                         ++
//++    -> disable receives and sends on socket                                             ++
//++    -> close socket                                                                     ++
//++                                                                                        ++
//++++++++++++++++++++++++++++++++++++++++++++++++++++++++++++++++++++++++++++++++++++++++++++

  case FSM_TCP of

    //**********************************************************************************
    _STATE_INIT_SERVER: // init state ... check if interface is present
    //**********************************************************************************
      if (bdStatus.ErrorNoUserInterface = true) then
        Control := _STATE_NO_USER_INTERFACE_CONNECTED;
      elsif (bdStatus.ErrAsyncTask = true) then
        Control := _STATE_ERROR_CREATING_TASK;
      elsif (bdStatus.ErrSema01 = true) | (bdStatus.ErrSema02 = true) then
        Control := _STATE_ERROR_CREATING_MUTEX;
      elsif (bdStatus.ErrMem = true) then
        Control := _STATE_ERROR_ALLOCATING_MEMORY;
      else
        if lsl_tcp_user <> NIL then
          FSM_TCP := _STATE_IDLE;
        else
          ErrorCode := -1;
        end_if;
      end_if;

    //**********************************************************************************
    _STATE_IDLE: // idle state ... wait for start server
    //**********************************************************************************
      FSM_TCP := _STATE_MAIN_SOCK;
      ActConn := 0;

    //**********************************************************************************
    _STATE_MAIN_SOCK: // allocate main socket
    //**********************************************************************************
      dMainSock := OS_TCP_USER_SOCKET();
      if (dMainSock < 0) then
        MainSocketError(FSM_TCP, TCP_SVR_ERR_GROUP_OS, dMainSock);
        FSM_TCP := _STATE_ERROR;
      else
        dRet := SetMainSocketOptions();
        if (dRet = TCP_SVR_NO_ERROR) then
          FSM_TCP := _STATE_LISTEN;
        else
          MainSocketError(FSM_TCP, TCP_SVR_ERR_GROUP_OS, dRet);
          ErrorCode := -12;
          FSM_TCP := _STATE_CLOSE_MAIN_SOCK;
        end_if;
      end_if;

    //**********************************************************************************
    _STATE_LISTEN: // listen for an incoming connection
    //**********************************************************************************
      dRet := OS_TCP_USER_LISTEN(dMainSock, to_UDINT(Port), to_udint(MaxConnections));
      if (dRet < 0) then
        if ((dRet = TCP_INVALID_SOCKET) | (dRet = TCP_INVALID_SOCKNUM)) then
          MainSocketError(FSM_TCP, TCP_SVR_ERR_GROUP_OS, dRet);
          FSM_TCP := _STATE_CLOSE_MAIN_SOCK;
        end_if;
      else
        FSM_TCP := _STATE_ACCEPT;
      end_if;

    //**********************************************************************************
    _STATE_ACCEPT: // accept a connection from any remote host
    //**********************************************************************************
      if (ActConn < MaxConn) then
        dNewSock := dAccSock := OS_TCP_USER_ACCEPT(dMainSock, 0);
        if (dAccSock < 0) & (dAccSock <> TCP_NOT_READY) then
          MainSocketError(FSM_TCP, TCP_SVR_ERR_GROUP_OS, dAccSock);
          FSM_TCP := _STATE_CLOSE_SOCK;
        elsif (dAccSock >= 0) then
          dRet := AddConnIntern(dAccSock, (#pConn)$^pVoid);
          if (dRet = TCP_SVR_NO_ERROR) & (pConn <> NIL) then
            dRet := SetSocketOptions(pConn);
            if (dRet = TCP_SVR_NO_ERROR) then
              FSM_TCP := _STATE_RECV;
              ErrorCode  := 0;
            else
              pConn^.FSM_TCP := _STATE_SHUTDOWN;
              ErrorCode := -12;
              FSM_TCP := _STATE_RECV;
            end_if;
          else
            FSM_TCP := _STATE_RECV;
          end_if;
        elsif (ActConn > 0) then
          FSM_TCP     := _STATE_RECV;
          ErrorCode      := 0;
        end_if;
      else
        FSM_TCP := _STATE_RECV;
      end_if;

    //**********************************************************************************
    _STATE_RECV: // general send and receive state
    //**********************************************************************************

      //loop to process more connections per run
      //i is not used, the pActConn will be advanced
      //if InhibNextConn is set (not all data of the current connection could be sent)
      //we stop the loop, and continue next run.
      if (ActConn < ConnectionsPerRun) then
        ConnPerRun := ActConn;
      else
        ConnPerRun := ConnectionsPerRun;
      end_if;
      for i := 1 to ConnPerRun do

        case pActConn^.FSM_TCP of

          (*===================================================================*)
          _STATE_RECV: // - RECEIVE DATA
          (*===================================================================*)
            dNewSock := pActConn^.dSocket;
            if (pActConn^.bdSettings.SockOptChanged = true) then
              pActConn^.FSM_TCP := _STATE_CONN_SOCK_OPT;
            else
              dBytes := OS_TCP_USER_NREAD_AVAILABLE(pActConn^.dSocket);
              if (dBytes <= 0) then
                if (dBytes <> TCP_NOT_READY) then
                  ConnSocketError(pActConn^.dSocket, pActConn^.FSM_TCP, TCP_SVR_ERR_GROUP_OS, dBytes);
                  pActConn^.FSM_TCP := _STATE_SHUTDOWN;
                  ErrorCode := -1;
                else
                  if (Timeout > 0) then
                    if ((ops.tAbsolute - pActConn^.udTimeStamp) > to_UDINT(Timeout)) then
                      ConnSocketError(pActConn^.dSocket, pActConn^.FSM_TCP, TCP_SVR_ERR_GROUP_AP, TCP_SVR_ERR_CODE_AP_TIMEOUT);
                      pActConn^.FSM_TCP := _STATE_SHUTDOWN;
                      ErrorCode := -2;
                    end_if;
                  end_if;
                end_if;

                pThisInterface^.DataHandling(dSocket:=pActConn^.dSocket, udAvailableData:=0);

              else
                if (dBytes > SizeOfTXBuffer$DINT) then
                  dBytes := SizeOfTXBuffer$DINT;
                end_if;

                UserDataToRead := pThisInterface^.DataHandling(dSocket:=pActConn^.dSocket, udAvailableData:=to_udint(dBytes));
                if UserDataToRead > to_udint(dBytes) then
                  UserDataToRead := to_udint(dBytes);
                end_if;

                if UserDataToRead > 0 then
                  dBytes := to_dint(UserDataToRead);
                  RECVbuffer.udSize := dBytes$UDINT;
                  dRet := OS_TCP_USER_RECV(pActConn^.dSocket, RECVbuffer.pData$^CHAR, dBytes$UDINT, 0, 0);
                  if (dRet = TCP_SOCK_NOT_CONNECTED) then
                    ConnSocketError(pActConn^.dSocket, pActConn^.FSM_TCP, TCP_SVR_ERR_GROUP_OS, dRet);
                    pActConn^.FSM_TCP := _STATE_SHUTDOWN;
                    ErrorCode := -3;
                  elsif (dRet <= 0) & (dRet <> TCP_NOT_READY) then
                    ConnSocketError(pActConn^.dSocket, pActConn^.FSM_TCP, TCP_SVR_ERR_GROUP_OS, dRet);
                    pActConn^.FSM_TCP := _STATE_SHUTDOWN;
                    ErrorCode := -1;
                  else
                    pThisInterface^.Response(RECVbuffer.pData, RECVbuffer.udSize, pActConn^.dSocket);
                    if (Timeout > 0) then
                      pActConn^.udTimeStamp := ops.tAbsolute;
                    end_if;
                  end_if;
                end_if;
              end_if;

              if (pActConn^.FSM_TCP = _STATE_RECV) then
                if pActConn^.BufferHeader.DataSize > 0 then
                  pActConn^.FSM_TCP := _STATE_SEND;
                elsif pActConn^.SendBuffer.udUsed > sizeof(_BUFFER_HEADER) then
                  pActConn^.pBufferWaitForSendingHelp := pActConn^.pBufferWaitForSendig;
                  pActConn^.FSM_TCP := _STATE_SEND;
                end_if;
              end_if;
            end_if;

          (*===================================================================*)
          _STATE_CONN_SOCK_OPT: // set socket options
          (*===================================================================*)
            dRet := SetSocketOptions(pActConn);
            if (dRet = TCP_SVR_NO_ERROR) then
              pActConn^.FSM_TCP := _STATE_RECV;
            else
              pActConn^.FSM_TCP := _STATE_SHUTDOWN;
            end_if;

          (*===================================================================*)
          _STATE_SEND:
          (*===================================================================*)
            if (ErrorCode <> -11) then
              if (pActConn^.BufferHeader.DataSize = 0) then
                dRet := RingbufferReadEntry(#pActConn^.SendBuffer, pActConn^.pBufferWaitForSendig, #pActConn^.BufferHeader.DataSize);
                pActConn^.pBufferWaitForSendingHelp := pActConn^.pBufferWaitForSendig;
              end_if;
              if (pActConn^.BufferHeader.DataSize > 0) then
                dRet := SendTCP(pActConn^.pBufferWaitForSendingHelp, pActConn^.BufferHeader.DataSize, pActConn^.dSocket, false);
                if (dRet >= 0) then
                  pActConn^.BufferHeader.DataSize -= dRet$UDINT;
                  pActConn^.pBufferWaitForSendingHelp += dRet;
                  if (pActConn^.BufferHeader.DataSize <= 0) then
                    pActConn^.FSM_TCP := _STATE_RECV;
                    pActConn^.pBufferWaitForSendingHelp := pActConn^.pBufferWaitForSendig;
                  else
                    bdStatus.InhibNextConn := true;
                  end_if;
                else
                  ConnSocketError(pActConn^.dSocket, pActConn^.FSM_TCP, TCP_SVR_ERR_GROUP_OS, dRet);
                  pActConn^.FSM_TCP := _STATE_RECV;
                  ErrorCode := -6;
                end_if;
              else
                pActConn^.FSM_TCP := _STATE_RECV;
              end_if;
            else
              pActConn^.FSM_TCP := _STATE_RECV;
            end_if;

          (*===================================================================*)
          _STATE_SHUTDOWN:
          (*===================================================================*)
            OS_TCP_USER_CLOSESOCKET(pActConn^.dSocket, pActConn^.CloseSocketType);
            pActConn^.FSM_TCP := _STATE_DEL_CONNECTION;

          (*===================================================================*)
          _STATE_DEL_CONNECTION:
          (*===================================================================*)
            DelConnIntern(pActConn^.dSocket);
            dNewSock := 0;

          (*===================================================================*)
          else // INAVLID CONNECTION STATE
          (*===================================================================*)
            pActConn^.FSM_TCP := _STATE_RECV;

        end_case;

        if (ActConn = 0) then
          exit;
        else
          if (bdStatus.InhibNextConn = false) then
            pActConn := pActConn^.pNextConn;
            if ((ops.tAbsolute - udTimeStamp) >= udTimeAccept) then
              FSM_TCP := _STATE_ACCEPT;
              udTimeStamp := ops.tAbsolute;
            end_if;
          else
            bdStatus.InhibNextConn := false;
            exit;
          end_if;
        end_if;

      end_for;

      if (ActConn = 0) then
        FSM_TCP := _STATE_ACCEPT;
      end_if;

    //**********************************************************************************
    _STATE_CLOSE_SOCK: // close all sockets
    //**********************************************************************************
      for i := 0 to (MaxConn-1) do
        if (SocketArray[i].dSocket <> 0) then
          OS_TCP_USER_CLOSESOCKET(SocketArray[i].dSocket, SocketArray[i].CloseSocketType);
          SocketArray[i].dSocket   := 0;
          SocketArray[i].FSM_TCP   := _STATE_IDLE;
          SocketArray[i].pNextConn := NIL;
        end_if;
      end_for;
      dNewSock := 0;
      ActConn := 0;
      FSM_TCP := _STATE_CLOSE_MAIN_SOCK;

    //**********************************************************************************
    _STATE_CLOSE_MAIN_SOCK: // close main socket
    //**********************************************************************************
        OS_TCP_USER_CLOSESOCKET(dMainSock, 0);
        dMainSock := 0;

        FSM_TCP := _STATE_IDLE;

    //**********************************************************************************
    _STATE_ERROR,
    _STATE_ERROR_ALLOCATING_MEMORY,
    _STATE_ERROR_CREATING_MUTEX,
    _STATE_ERROR_CREATING_TASK,
    _STATE_NO_USER_INTERFACE_CONNECTED:
    //**********************************************************************************

  end_case;

//+++++++++++++++++++++++++++++++++++++++++++++++++++++++++++++++++++++++++++++++++++++++++++
//++                                       E N D                                           ++
//+++++++++++++++++++++++++++++++++++++++++++++++++++++++++++++++++++++++++++++++++++++++++++

  Control := FSM_TCP;

END_FUNCTION

FUNCTION _TCPIPServer::SendTCP
	VAR_INPUT
		pData 	: ^void;
		udSize 	: UDINT;
		dSock 	: DINT;
		bDirect 	: DINT;
	END_VAR
	VAR_OUTPUT
		dRetcode 	: DINT;
	END_VAR

  if ((FSM_TCP <> _STATE_RECV) & (bDirect = false)) then
    dRetcode := -1;
    return;
  end_if;

  dRetcode := OS_TCP_USER_SEND(dSock, pData$^CHAR, udSize, 0, 0);

END_FUNCTION

FUNCTION _TCPIPServer::SENDbuffer_Read
	VAR_INPUT
		pBuffer 	: ^_TX_RINGBUFFER;
		pData 	: ^void;
		udSize 	: UDINT;
	END_VAR
	VAR_OUTPUT
		Retcode 	: DINT;
	END_VAR
VAR
	udBytes2End   : UDINT;
  udBytesTmp    : UDINT;
END_VAR

  Retcode := 0;

  if (pBuffer = NIL) | (pData = NIL) | (pBuffer^.pMem = NIL) then
    return; //### invalid pointer
  end_if;

  udBytes2End := (pBuffer^.pMem$UDINT + pBuffer^.udSize) - pBuffer^.pRead$UDINT;

  if (udSize > udBytes2End) then

    //##########################################################################################
    //### we must read the data in 2 blocks (|second|...........other data...........|first|)
    //##########################################################################################
    _memcpy(ptr1 := pData, ptr2 := pBuffer^.pRead, cntr := udBytes2End); //### copy the first block
    pData += udBytes2End;
    pBuffer^.pRead := pBuffer^.pMem$^USINT;
    udBytesTmp := udSize - udBytes2End;
    _memcpy(ptr1 := pData, ptr2 := pBuffer^.pRead, cntr := udBytesTmp); //### copy the second block
    pBuffer^.pRead += udBytesTmp;

  else

    //##########################################################################################
    //### read data in one block
    //##########################################################################################
    _memcpy(ptr1 := pData, ptr2 := pBuffer^.pRead, cntr := udSize);
    pBuffer^.pRead += udSize;
  end_if;

  pBuffer^.udUsed -= udSize; // decrease the number of bytes in ringbuffer
  Retcode := udSize$DINT;

END_FUNCTION

FUNCTION _TCPIPServer::SENDbuffer_Write
	VAR_INPUT
		pData 	: ^void;
		udSize 	: UDINT;
		pBuffer 	: ^_TX_RINGBUFFER;
	END_VAR
	VAR_OUTPUT
		dRetcode 	: DINT;
	END_VAR
VAR
	udBytes2End   : UDINT;
  udBytesTmp    : UDINT;
END_VAR

  if (pBuffer^.pMem = NIL) | (pData = NIL) | (pBuffer = NIL) then         // Check if Pointer is NIL
    dRetcode := -9;                       // Pointer to SendBuffer is NIL
    return;
  end_if;

  dRetcode := 0;

  if ((udSize) > (pBuffer^.udSize - pBuffer^.udUsed)) then
    return; //### buffer full
  end_if;

  udBytes2End := (pBuffer^.pMem$UDINT + pBuffer^.udSize) - pBuffer^.pWrite$UDINT; // calculate number of bytes till the end of SENDbuffer

  if (udSize > udBytes2End) then

    //##########################################################################################
    //### we must write the data in 2 blocks  (|second|...........other data...........|first|)
    //##########################################################################################
    _memcpy(ptr1 := pBuffer^.pWrite, ptr2 := pData, cntr := udBytes2End); // copy the first block
    pData += udBytes2End;
    pBuffer^.pWrite := pBuffer^.pMem$^USINT;
    udBytesTmp := udSize - udBytes2End;
    _memcpy(ptr1 := pBuffer^.pWrite, ptr2 := pData, cntr := udBytesTmp); // copy the second block
    pBuffer^.pWrite += udBytesTmp;
    dRetcode := udSize$DINT;
  else

    //##########################################################################################
    //### store data in one block
    //##########################################################################################
    _memcpy(ptr1 := pBuffer^.pWrite, ptr2 := pData, cntr := udSize);
    pBuffer^.pWrite += udSize;
    dRetcode := udSize$DINT;
  end_if;

  pBuffer^.udUsed += udSize; // increase the number of bytes in ringbuffer

END_FUNCTION

FUNCTION VIRTUAL GLOBAL _TCPIPServer::SendData
	VAR_INPUT
		pData 	: ^void;
		udSize 	: UDINT;
		dSock 	: DINT;
		bDirect 	: BOOL;
	END_VAR
	VAR_OUTPUT
		dRetcode 	: DINT;
	END_VAR
VAR
  dRet        : DINT;
  i           : USINT;
  bFound      : BOOL;
END_VAR

  if (bDirect = true) then
    if (udSize <= 1452) then
      dRet := SendTCP(pData, udSize, dSock, true);
      if (dRet <> udSize$DINT) then
        dRetcode := -6;
      else
        dRetcode := dRet;
      end_if;
    else
      dRetcode := -13;
      ErrorCode   := -13;
    end_if;
  else

    bFound := false;
    for i := 0 to (MaxConn-1)$USINT do
      if (SocketArray[i].dSocket = dSock) then
        bFound := true;
        exit;
      end_if;
    end_for;

    if (bFound = true) then
      dRet := RingbufferWriteEntry(#SocketArray[i].SendBuffer, pData, udSize);
      if (dRet = TCP_SVR_NO_ERROR) then
        dRetcode := to_DINT(udSize);
      else
        dRetcode := -11;
        ErrorCode   := -11;
      end_if;
    else
      dRetcode := -11;
      ErrorCode   := -11;
    end_if;

  end_if;

END_FUNCTION

FUNCTION _TCPIPServer::Read_LSLOBJ_CRC32
	VAR_INPUT
		pCRC32 	: ^CHAR;
	END_VAR
	VAR_OUTPUT
		Retcode 	: DINT;
	END_VAR
VAR
	udStrLen    : UDINT;
  udCRC32     : UDINT;
  szObjName   : ARRAY [0..255] OF CHAR;
END_VAR

  Retcode := TCP_SVR_NO_ERROR;

  if (pCRC32 <> NIL) then
    pCRC32^ := 0x00;
    udStrLen := _GetObjName(this, #szObjName[0]);
    if (udStrLen > 0) then
      udCRC32 := CheckSum.CRC32(#szObjName[0], udStrLen, 0);
      SigCLib.IToA(udCRC32$DINT, pCRC32, 0x10);
    else
      Retcode := TCP_SVR_ERR_GET_LSLOBJ_NAME;
    end_if;
  else
    Retcode := TCP_SVR_ERR_INVALID_POINTER;
  end_if;

END_FUNCTION

FUNCTION _TCPIPServer::Read_AP_TaskPeriod
	VAR_OUTPUT
		Retcode 	: DINT;
	END_VAR
VAR
	dRet          : DINT;
  LSLOBJ_INFO   : LSLOBJ_INFO;
END_VAR

  Retcode := TCP_SVR_NO_ERROR;

  dRet := _TaskObjectControl.GetObjectInfo(this, OBJ_CT, #LSLOBJ_INFO);
  case dRet of
    (*=============================================================================*)
    0: // - GET OBJECT INFO OK
    (*=============================================================================*)
      if (bdStatus.SalamanderOS = true) then
        // --------------------------------------------------------
        // - SALAMANDER OS
        // --------------------------------------------------------
        if (LSLOBJ_INFO.orgperiod AND 0x80000000) then
          // -------------------------------------------------------
          // - TASK PERIOD IN [µs]
          // -------------------------------------------------------
          AP_TaskTime  := LSLOBJ_INFO.orgperiod XOR 0x80000000;
        else
          // -------------------------------------------------------
          // - TASK PERIOD IN [ms]
          // -------------------------------------------------------
          AP_TaskTime  := LSLOBJ_INFO.orgperiod * 1000;
        end_if;
      else
        // --------------------------------------------------------
        // - LASAL OS
        // --------------------------------------------------------
        if (LSLOBJ_INFO.orgperiod AND 0x80000000) then
          // -------------------------------------------------------
          // - TASK PERIOD IN [µs]
          // -------------------------------------------------------
          AP_TaskTime := (LSLOBJ_INFO.orgperiod XOR 0x80000000) / 1000;
          if (AP_TaskTime = 0) then
            AP_TaskTime := 1;
          end_if;
        else
          // -------------------------------------------------------
          // - TASK PERIOD IN [ms]
          // -------------------------------------------------------
          AP_TaskTime  := LSLOBJ_INFO.orgperiod;
        end_if;
      end_if;

    (*=============================================================================*)
    -1: // - ERROR READ OBJECT INFO (NO APPLICATION)
    (*=============================================================================*)
      Retcode     := TCP_SVR_ERR_TASK_TIME_NO_APP;
      AP_TaskTime := 0xFFFFFFFF;

    (*=============================================================================*)
    -3: // - ERROR READ OBJECT INFO (NO APPLICATION)
    (*=============================================================================*)
      Retcode     := TCP_SVR_ERR_TASK_TIME_WRONG_TASK_TYPE;
      AP_TaskTime := 0xFFFFFFFF;

    (*=============================================================================*)
    -5: // - OBJECT NOT FOUND (TASK DEACTIVATED)
    (*=============================================================================*)
      Retcode     := TCP_SVR_ERR_TASK_TIME_OBJ_NOT_FOUND;
      AP_TaskTime := 0xFFFFFFFF;

  end_case;

END_FUNCTION

FUNCTION _TCPIPServer::AP_TaskCreate
	VAR_INPUT
		pTaskName 	: ^CHAR;
		pCallback 	: ^void;
	END_VAR
	VAR_OUTPUT
		Retcode 	: DINT;
	END_VAR

  Retcode := TCP_SVR_NO_ERROR;

  AP_TaskHandle := _MultiTask.CREATETHREAD(pCallback, AP_TaskPriority, 0x4000, MT_TASK_SAVETHIS, this, pTaskName);
  if (AP_TaskHandle = NIL) then
    Retcode := TCP_SVR_ERR_TASK_CREATE;
  end_if;

END_FUNCTION

FUNCTION _TCPIPServer::AP_TaskCallback
	VAR_INPUT
		Param0 	: ^void;
	END_VAR

  while 1 do
    CyclicCall();
    AP_TaskDelay(AP_TaskTime);
  end_while;

END_FUNCTION

FUNCTION _TCPIPServer::GetMultiTaskErrorCode
	VAR_INPUT
		pErrTxt 	: ^CHAR;
	END_VAR
VAR
	ErrMT     : DINT;
END_VAR

  ErrMT := _MultiTask.GETLASTERROR();
  case ErrMT of

    (*===============================================================================================*)
    MTERROR_NONE: // - NO ERROR
    (*===============================================================================================*)
      SigCLib.StrCpy(pErrTxt, "MTERROR_NONE");

    (*===============================================================================================*)
    MTERROR_NOMEM: // - NO MORE MEMORY TO RUN THIS FUNCTION, E.G. INTERNAL ALLOC FAILED
    (*===============================================================================================*)
      SigCLib.StrCpy(pErrTxt, "MTERROR_NOMEM");

    (*===============================================================================================*)
    MTERROR_NOFCT: // - CREATE TASK NEEDS A VALID TASK FUNCTION
    (*===============================================================================================*)
      SigCLib.StrCpy(pErrTxt, "MTERROR_NOFCT");

    (*===============================================================================================*)
    MTERROR_FCTNOTINMEM: // - CREATE TASK NEEDS A TASK FUNCTION PLACED IN LASAL CODE MEMORY
    (*===============================================================================================*)
      SigCLib.StrCpy(pErrTxt, "MTERROR_FCTNOTINMEM");

    (*===============================================================================================*)
    MTERROR_WRONGPRIOR: // - CREATE TASK ONLY SUPPORTS PRIORS FROM 1 .. 14
    (*===============================================================================================*)
      SigCLib.StrCpy(pErrTxt, "MTERROR_WRONGPRIOR");

    (*===============================================================================================*)
    MTERROR_STACK: // - CREATE TASK ONLY SUPPORT SATCK SIZE LOWER THAN 0x4000
    (*===============================================================================================*)
      SigCLib.StrCpy(pErrTxt, "MTERROR_STACK");

    (*===============================================================================================*)
    MTERROR_NAME: // - CREATE TASK, MAILBOX OR SEMAPHORE NEEDS A VALID NAME
    (*===============================================================================================*)
      SigCLib.StrCpy(pErrTxt, "MTERROR_NAME");

    (*===============================================================================================*)
    MTERROR_NAMEUSED: // - CREATE TASK, MAILBOX OR SEMAPHORE NAME ALREADY IN USE
    (*===============================================================================================*)
      SigCLib.StrCpy(pErrTxt, "MTERROR_NAMEUSED");

    (*===============================================================================================*)
    MTERROR_HANDLE: // - HANDLE NOT FOUND IN OS-LIST => NOT VALID
    (*===============================================================================================*)
      SigCLib.StrCpy(pErrTxt, "MTERROR_HANDLE");

    (*===============================================================================================*)
    MTERROR_NOTALLOWED: // - MT-FUNCTION NOT ALLOWED IN THIS TASK CONTEXT
    (*===============================================================================================*)
      SigCLib.StrCpy(pErrTxt, "MTERROR_NOTALLOWED");

    (*===============================================================================================*)
    MTERROR_MESSAGESIZE: // - MAILBOX NEED A VALID MESSAGE SIZE
    (*===============================================================================================*)
      SigCLib.StrCpy(pErrTxt, "MTERROR_MESSAGESIZE");

    (*===============================================================================================*)
    MTERROR_DATA: // - POINTER TO DATA IS NOT VALID
    (*===============================================================================================*)
      SigCLib.StrCpy(pErrTxt, "MTERROR_DATA");

    (*===============================================================================================*)
    MTERROR_PTR: // - INVALID POINTER, PARAMETER OR INTERNAL
    (*===============================================================================================*)
      SigCLib.StrCpy(pErrTxt, "MTERROR_PTR");

    (*===============================================================================================*)
    MTERROR_TASKID: // - INVALID TASK ID, ID NOT FOUND
    (*===============================================================================================*)
      SigCLib.StrCpy(pErrTxt, "MTERROR_TASKID");

    (*===============================================================================================*)
    MTERROR_NOTASK: // - TASK DOES NOT EXIST
    (*===============================================================================================*)
      SigCLib.StrCpy(pErrTxt, "MTERROR_NOTASK");

    (*===============================================================================================*)
    MTERROR_NOIFFNC: // - INTERFACE FUNCTION IS NOT AVAILABLE
    (*===============================================================================================*)
      SigCLib.StrCpy(pErrTxt, "MTERROR_NOIFFNC");

    (*===============================================================================================*)
    else // - UNKNOWN ERROR CODE
    (*===============================================================================================*)
      SigCLib.StrCpy(pErrTxt, "MTERROR_UNKNOWN");

  end_case;

END_FUNCTION

FUNCTION _TCPIPServer::AP_SemaCreate
	VAR_INPUT
		pSemaName 	: ^CHAR;
		Index 	: DINT;
	END_VAR
	VAR_OUTPUT
		Retcode 	: DINT;
	END_VAR

  Retcode := TCP_SVR_NO_ERROR;

  if (pSemaName <> NIL) then
    case Index of
      (*=================================================================================*)
      0:
      (*=================================================================================*)
        AP_SemaHandle1 := _MultiTask.CREATESEMAPHORE(MTSEMATYPE_MUTEX, 1, 0, pSemaName);
        if (AP_SemaHandle1 = NIL) then
          Retcode := TCP_SVR_ERR_SEMA_CREATE;
        end_if;

      (*=================================================================================*)
      1:
      (*=================================================================================*)
        AP_SemaSockOpt := _MultiTask.CREATESEMAPHORE(MTSEMATYPE_MUTEX, 1, 0, pSemaName);
        if (AP_SemaSockOpt = NIL) then
          Retcode := TCP_SVR_ERR_SEMA_CREATE;
        end_if;

      (*=================================================================================*)
      else
      (*=================================================================================*)
        Retcode := TCP_SVR_ERR_SEMA_INVALID_IDX;

    end_case;
  else
    Retcode := TCP_SVR_ERR_SEMA_INVALID_NAME;
  end_if;

END_FUNCTION

FUNCTION _TCPIPServer::AP_TaskDelay
	VAR_INPUT
		udTaskDelay 	: UDINT;
	END_VAR

  if (bdStatus.SalamanderOS = true) then
    OSSD_DELAY(pCIL_DEBUG, udTaskDelay);
  else
    _MultiTask.TASKDELAY(udTaskDelay);
  end_if;

END_FUNCTION

FUNCTION _TCPIPServer::SetMainSocketOptions
	VAR_OUTPUT
		Retcode 	: DINT;
	END_VAR
VAR
	dRet        : DINT;
  OptionValue : DINT;
END_VAR

  Retcode := TCP_SVR_NO_ERROR;

  OptionValue := 1;
  dRet := OS_TCP_USER_SETSOCKOPT(dMainSock, SOL_SOCKET, SO_REUSEADDR, #OptionValue$CHAR, sizeof(DINT));
  if (dRet <> 0) then
    Retcode := dRet;
  end_if;

  OptionValue := 0;
  dRet := OS_TCP_USER_SETSOCKOPT(dMainSock, SOL_SOCKET, SO_DELAYED_ACK, #OptionValue$CHAR, sizeof(DINT));
  if (dRet <> 0) then
    Retcode := dRet;
  end_if;

END_FUNCTION

FUNCTION _TCPIPServer::RingbufferReadEntry
	VAR_INPUT
		pBuffer 	: ^_TX_RINGBUFFER;
		pData 	: ^void;
		pSize 	: ^UDINT;
	END_VAR
	VAR_OUTPUT
		Retcode 	: DINT;
	END_VAR
VAR
	BufferHeader    : _BUFFER_HEADER;
  dRet            : DINT;
END_VAR

  Retcode := TCP_SVR_NO_ERROR;
  pSize^  := 0;

  if (pBuffer = NIL) | (pData = NIL) | (pSize = NIL) then
    Retcode := TCP_SVR_ERR_INVALID_POINTER;
  else
    if (pBuffer^.udUsed = 0) then
      Retcode := TCP_SVR_SEND_BUFFER_EMPTY;
    else
      AP_SemaWait(AP_SemaHandle1);
      dRet := SENDBuffer_Read(pBuffer, #BufferHeader, sizeof(_BUFFER_HEADER));
      if (dRet = sizeof(_BUFFER_HEADER)) then
        dRet := SENDBuffer_Read(pBuffer, pData, BufferHeader.DataSize);
        if (dRet = BufferHeader.DataSize$DINT) then
          pSize^ := BufferHeader.DataSize;
        else
          Retcode := TCP_SVR_ERR_SEND_BUFFER_FATAL_ERROR;
        end_if;
      else
        Retcode := TCP_SVR_ERR_SEND_BUFFER_FATAL_ERROR;
      end_if;
      AP_SemaSignal(AP_SemaHandle1);
    end_if;
  end_if;

END_FUNCTION

FUNCTION _TCPIPServer::RingbufferWriteEntry
	VAR_INPUT
		pBuffer 	: ^_TX_RINGBUFFER;
		pData 	: ^void;
		udSize 	: UDINT;
	END_VAR
	VAR_OUTPUT
		Retcode 	: DINT;
	END_VAR
VAR
	BufferHeader  : _BUFFER_HEADER;
END_VAR

  Retcode := TCP_SVR_NO_ERROR;

  if (pBuffer = NIL) | (pData = NIL) then
    Retcode := TCP_SVR_ERR_INVALID_POINTER;
  else
    AP_SemaWait(AP_SemaHandle1);
    if ((udSize + sizeof(_BUFFER_HEADER)) > (pBuffer^.udSize - pBuffer^.udUsed)) then
      Retcode := TCP_SVR_SEND_BUFFER_FULL;
    else
      BufferHeader.DataSize := udSize;
      SENDbuffer_Write(#BufferHeader, sizeof(_BUFFER_HEADER), pBuffer);
      SENDbuffer_Write(pData, udSize, pBuffer);
    end_if;
    AP_SemaSignal(AP_SemaHandle1);
  end_if;

END_FUNCTION

FUNCTION _TCPIPServer::AP_SemaWait
	VAR_INPUT
		SemaHandle 	: MT_SEMAHANDLE;
	END_VAR

  if (SemaHandle <> NIL) then
    _MultiTask.WAIT(SemaHandle);
  end_if;

END_FUNCTION

FUNCTION _TCPIPServer::AP_SemaSignal
	VAR_INPUT
		SemaHandle 	: MT_SEMAHANDLE;
	END_VAR

  if (SemaHandle <> NIL) then
    _MultiTask.SIGNAL(SemaHandle);
  end_if;

END_FUNCTION

FUNCTION _TCPIPServer::SetSocketOptions
	VAR_INPUT
		pConn 	: ^_CONNECTION;
	END_VAR
	VAR_OUTPUT
		Retcode 	: DINT;
	END_VAR
VAR
	OptionValue       : DINT;
  dRet              : DINT;
  KeepAliveLasalOS  : _KeepAliveParaLasalOS;
END_VAR

  Retcode := TCP_SVR_NO_ERROR;

  AP_SemaWait(AP_SemaSockOpt);

  // -----------------------------------------------------------
  // - SOCKET OPTION NAGLE
  // -----------------------------------------------------------
  if (pConn^.ConnSockOpt.Nagle = true) then
    OptionValue := 1;
  else
    OptionValue := 0;
  end_if;
  dRet := OS_TCP_USER_SETSOCKOPT(pConn^.dSocket, SOL_SOCKET, SO_NAGLE, (#OptionValue)$^CHAR, sizeof(DINT));
  if (dRet < 0) then
    Retcode := dRet;
    ConnSocketError(pConn^.dSocket, pConn^.FSM_TCP, TCP_SVR_ERR_GROUP_OS, dRet);
  end_if;

  // -----------------------------------------------------------
  // - SOCKET OPTION KEEP ALIVE
  // -----------------------------------------------------------
  if (bdStatus.SalamanderOS = false) then
    // --------------------------------------------------------
    // - LASAL OS
    // --------------------------------------------------------
    if (pConn^.ConnSockOpt.KeepAlive = true) then
      KeepAliveLasalOS.interval := to_UINT(pConn^.KeepAlivePara.keepIDLE);
      KeepAliveLasalOS.retry    := to_UINT(pConn^.KeepAlivePara.keepINTVL);
      KeepAliveLasalOS.timeout  := to_UINT(pConn^.KeepAlivePara.keepCNT * pConn^.KeepAlivePara.keepINTVL);
    else
      KeepAliveLasalOS.interval := 0;
      KeepAliveLasalOS.retry    := 0;
      KeepAliveLasalOS.timeout  := 0;
    end_if;
    dRet := OS_TCP_USER_SETSOCKOPT(pConn^.dSocket, SOL_SOCKET, 8, (#KeepAliveLasalOS)$^CHAR, sizeof(_KeepAliveParaLasalOS));
    if (dRet < 0) then
      Retcode := dRet;
      ConnSocketError(pConn^.dSocket, pConn^.FSM_TCP, TCP_SVR_ERR_GROUP_OS, dRet);
    end_if;
  else
    // --------------------------------------------------------
    // - SALAMANDER OS
    // --------------------------------------------------------
    if (pConn^.ConnSockOpt.KeepAlive = true) then
      OptionValue := 1;
    else
      OptionValue := 0;
    end_if;
    dRet := OS_TCP_USER_SETSOCKOPT(pConn^.dSocket, SOL_SOCKET, 8, (#OptionValue)$^CHAR, sizeof(DINT));
    if (dRet < 0) then
      Retcode := dRet;
      ConnSocketError(pConn^.dSocket, pConn^.FSM_TCP, TCP_SVR_ERR_GROUP_OS, dRet);
    end_if;

//    if (pConn^.ConnSockOpt.KeepAlive = true) then
//      OptionValue := KeepAlivePara.keepCNT;
//      dRet := OS_TCP_USER_SETSOCKOPT(pConn^.dSocket, SOL_TCP, TCP_KEEPCNT, (#OptionValue)$^CHAR, sizeof(DINT));
//      if (dRet < 0) then
//        Retcode := dRet;
//        ConnSocketError(pConn^.dSocket, pConn^.FSM_TCP, TCP_SVR_ERR_GROUP_OS, dRet);
//      end_if;
//      OptionValue := KeepAlivePara.keepIDLE;
//      dRet := OS_TCP_USER_SETSOCKOPT(pConn^.dSocket, SOL_TCP, TCP_KEEPIDLE, (#OptionValue)$^CHAR, sizeof(DINT));
//      if (dRet < 0) then
//        Retcode := dRet;
//        ConnSocketError(pConn^.dSocket, pConn^.FSM_TCP, TCP_SVR_ERR_GROUP_OS, dRet);
//      end_if;
//      OptionValue := KeepAlivePara.keepINTVL;
//      dRet := OS_TCP_USER_SETSOCKOPT(pConn^.dSocket, SOL_TCP, TCP_KEEPINTVL, (#OptionValue)$^CHAR, sizeof(DINT));
//      if (dRet < 0) then
//        Retcode := dRet;
//        ConnSocketError(pConn^.dSocket, pConn^.FSM_TCP, TCP_SVR_ERR_GROUP_OS, dRet);
//      end_if;
//    end_if;
  end_if;

  // -----------------------------------------------------------
  // - SOCKET OPTION DELAYED ACK
  // -----------------------------------------------------------
  if (pConn^.ConnSockOpt.DelayedAck = true) then
    OptionValue := 1;
  else
    OptionValue := 0;
  end_if;
  OS_TCP_USER_SETSOCKOPT(pConn^.dSocket, SOL_SOCKET, SO_DELAYED_ACK, (#OptionValue)$^CHAR, sizeof(DINT));
  if (dRet < 0) then
    Retcode := dRet;
    ConnSocketError(pConn^.dSocket, pConn^.FSM_TCP, TCP_SVR_ERR_GROUP_OS, dRet);
  end_if;

  // -----------------------------------------------------------
  // - SOCKET OPTION REUSE ADDR
  // -----------------------------------------------------------
  if (pConn^.ConnSockOpt.ReuseAddr = true) then
    OptionValue := 1;
  else
    OptionValue := 0;
  end_if;
  OS_TCP_USER_SETSOCKOPT(pConn^.dSocket, SOL_SOCKET, SO_REUSEADDR, (#OptionValue)$^CHAR, sizeof(DINT));
  if (dRet < 0) then
    Retcode := dRet;
    ConnSocketError(pConn^.dSocket, pConn^.FSM_TCP, TCP_SVR_ERR_GROUP_OS, dRet);
  end_if;

  pConn^.bdSettings.SockOptChanged := false;

  AP_SemaSignal(AP_SemaSockOpt);

END_FUNCTION

FUNCTION _TCPIPServer::AddConnIntern
	VAR_INPUT
		dSocket 	: DINT;
		ppConn 	: ^pVoid;
	END_VAR
	VAR_OUTPUT
		Retcode 	: DINT;
	END_VAR
VAR
	i           : USINT;
  pFirstConn  : ^_CONNECTION;
  pNewConn    : ^_CONNECTION;
  pSearchConn : ^_CONNECTION;
END_VAR

  Retcode := TCP_SVR_NO_ERROR;
  if (ppConn <> NIL) then
    ppConn^ := NIL;
  end_if;

  if (ActConn < MaxConn) then

    for i := 0 to (MaxConn-1) do
      pFirstConn := #SocketArray[0] + (i * sizeof(_CONNECTION));
      if (pFirstConn^.dSocket <> 0) then
        exit;
      else
        pFirstConn := NIL;
      end_if;
    end_for;

    for i := 0 to (MaxConn-1) do
      pNewConn := #SocketArray[0] + (i * sizeof(_CONNECTION));
      if (pNewConn^.dSocket = 0) then
        pNewConn^.dSocket         := dSocket;
        pNewConn^.FSM_TCP         := _STATE_RECV;
        pNewConn^.ConnSockOpt     := MainSockOpt;
        pNewConn^.KeepAlivePara   := KeepAlivePara;
        pNewConn^.CloseSocketType := CloseSocketType;
        pNewConn^.bdSettings.SockOptChanged := true;
        ConnSocketInfo(dSocket, TCP_SVR_SOCK_INFO_CONNECT, 0);
        if (ppConn <> NIL) then
          ppConn^$^_CONNECTION := pNewConn;
        end_if;
        exit;
      end_if;
    end_for;

    if (pFirstConn = NIL) then
      pNewConn^.pNextConn := pNewConn;
    else
      pSearchConn := pFirstConn;
      while (pSearchConn^.pNextConn <> pFirstConn) do
        pSearchConn := pSearchConn^.pNextConn;
      end_while;
      pNewConn^.pNextConn    := pFirstConn;
      pSearchConn^.pNextConn := pNewConn;
    end_if;

    ActConn += 1;
    if (ActConn = 1) then
      pActConn := pNewConn;
    end_if;

    if (Timeout > 0) then
      pNewConn^.udTimeStamp := ops.tAbsolute;
    end_if;

  else
    Retcode := TCP_SVR_ERR_MAX_CONN;
  end_if;

END_FUNCTION

FUNCTION _TCPIPServer::DelConnIntern
	VAR_INPUT
		dSocket 	: DINT;
	END_VAR
	VAR_OUTPUT
		Retcode 	: DINT;
	END_VAR
VAR
	pConn       : ^_CONNECTION;
  pSearchConn : ^_CONNECTION;
  i           : USINT;
END_VAR

  Retcode := TCP_SVR_NO_ERROR;

  if (ActConn > 0) then

    for i := 0 to (MaxConn-1) do
      pConn := #SocketArray[0] + (i * sizeof(_CONNECTION));
      if (pConn^.dSocket = dSocket) then
        exit;
      else
        pConn := NIL;
      end_if;
    end_for;

    if (pConn <> NIL) then
      if (pConn^.pNextConn = pConn) then
        // - ONE ACTIVE CONNECTION
      else
        pSearchConn := pConn;
        while (pSearchConn^.pNextConn <> pConn) do
          pSearchConn := pSearchConn^.pNextConn;
        end_while;
        pSearchConn^.pNextConn := pConn^.pNextConn;
        pActConn := pConn^.pNextConn;
        bdStatus.InhibNextConn := true;
      end_if;
      pConn^.dSocket   := 0;
      pConn^.FSM_TCP   := _STATE_IDLE;
      pConn^.pNextConn := NIL;
      ConnSocketInfo(dSocket, TCP_SVR_SOCK_INFO_DISCONNECT, 0);
      ActConn -= 1;
    end_if;

  else
    // - ERROR NO CONN
  end_if;

END_FUNCTION

FUNCTION _TCPIPServer::ConnSocketInfo
	VAR_INPUT
		dSock 	: DINT;
		InfoPara1 	: DINT;
		InfoPara2 	: DINT;
	END_VAR

  if pThisInterface <> NIL then
    pThisInterface^.ConnSocketInfo(dSock, InfoPara1, InfoPara2);
  end_if;

END_FUNCTION

FUNCTION _TCPIPServer::ConnSocketError
	VAR_INPUT
		dSock 	: DINT;
		FSM_TCP 	: _FSM_TCPIP_SERVER;
		ErrGroup 	: DINT;
		ErrCode 	: DINT;
	END_VAR

  if pThisInterface <> NIL then
    pThisInterface^.ConnSocketError(dSock, FSM_TCP, ErrGroup, ErrCode);
  end_if;

END_FUNCTION

FUNCTION _TCPIPServer::MainSocketError
	VAR_INPUT
		FSM_TCP 	: _FSM_TCPIP_SERVER;
		ErrGroup 	: DINT;
		ErrCode 	: DINT;
	END_VAR

  if pThisInterface <> NIL then
    pThisInterface^.MainSocketError(FSM_TCP, ErrGroup, ErrCode);
  end_if;

END_FUNCTION

FUNCTION VIRTUAL GLOBAL _TCPIPServer::SetMainParameter
	VAR_INPUT
		Cmd 	: DINT;
		SubCmd 	: DINT;
		ParaValue 	: DINT;
	END_VAR
	VAR_OUTPUT
		Retcode 	: DINT;
	END_VAR

  Retcode := TCP_SVR_NO_ERROR;

  if (usInit > 0) then
    case Cmd of
      (*================================================================*)
      SVR_TCP_CMD_SETSOCKOPT:
      (*================================================================*)
        case SubCmd of
          (*==================================================*)
          SVR_TCP_SOCKOPT_NAGLE:
          (*==================================================*)
            if (ParaValue = 0) then
              MainSockOpt.Nagle := false;
            else
              MainSockOpt.Nagle := true;
            end_if;
          (*==================================================*)
          SVR_TCP_SOCKOPT_KEEPALIVE:
          (*==================================================*)
            if (ParaValue = 0) then
              MainSockOpt.KeepAlive := false;
            else
              MainSockOpt.KeepAlive := true;
            end_if;
          (*==================================================*)
          SVR_TCP_SOCKOPT_DELAYEDACK:
          (*==================================================*)
            if (ParaValue = 0) then
              MainSockOpt.DelayedAck := false;
            else
              MainSockOpt.DelayedAck := true;
            end_if;
          (*==================================================*)
          SVR_TCP_SOCKOPT_REUSEADDR:
          (*==================================================*)
            if (ParaValue = 0) then
              MainSockOpt.ReuseAddr := false;
            else
              MainSockOpt.ReuseAddr := true;
            end_if;
          (*==================================================*)
          else // - INVALID SUB COMMAND
          (*==================================================*)
            Retcode := TCP_SVR_ERR_SET_PARA_INVALID_SUB_CMD;
        end_case;

      (*================================================================*)
      SVR_TCP_CMD_TASKPRIO: // - ASYNC TASK PRIORITY
      (*================================================================*)
        case SubCmd of
          (*==================================================*)
          SVR_TCP_SUB_CMD_TASKPRIO:
          (*==================================================*)
            if (usInit < INIT_FIRSTSCAN) then
              AP_TaskPriority := ParaValue$UDINT;
            else
              Retcode := TCP_SVR_ERR_TASK_ALREADY_EXIST;
            end_if;
          (*==================================================*)
          else // - INVALID SUB COMMAND
          (*==================================================*)
            Retcode := TCP_SVR_ERR_SET_PARA_INVALID_SUB_CMD;
        end_case;

      (*================================================================*)
      SVR_TCP_CMD_KEEPALIVEPARA: // - ASYNC TASK PRIORITY
      (*================================================================*)
        case SubCmd of
          (*==================================================*)
          SVR_TCP_KEEPALIVE_KEEPIDLE:
          (*==================================================*)
            KeepAlivePara.keepIDLE := ParaValue;
          (*==================================================*)
          SVR_TCP_KEEPALIVE_KEEPINTVL:
          (*==================================================*)
            KeepAlivePara.keepINTVL := ParaValue;
          (*==================================================*)
          SVR_TCP_KEEPALIVE_KEEPCNT:
          (*==================================================*)
            KeepAlivePara.keepCNT := ParaValue;
          (*==================================================*)
          else // - INVALID SUB COMMAND
          (*==================================================*)
            Retcode := TCP_SVR_ERR_SET_PARA_INVALID_SUB_CMD;
        end_case;

      (*================================================================*)
      SVR_TCP_CMD_CLOSESOCKETTYPE:
      (*================================================================*)
        case SubCmd of
          (*==================================================*)
          SVR_TCP_CLOSESOCKETTYPE:
          (*==================================================*)
            CloseSocketType := ParaValue$UDINT;
          (*==================================================*)
          else // - INVALID SUB COMMAND
          (*==================================================*)
            Retcode := TCP_SVR_ERR_SET_PARA_INVALID_SUB_CMD;
        end_case;

      (*================================================================*)
      else // - INVALID COMMAND
      (*================================================================*)
        Retcode := TCP_SVR_ERR_SET_PARA_INVALID_CMD;

    end_case;
  else
    Retcode := TCP_SVR_ERR_MAIN_INIT;
  end_if;

END_FUNCTION

FUNCTION VIRTUAL GLOBAL _TCPIPServer::SetSocketParameter
	VAR_INPUT
		dSock 	: DINT;
		Cmd 	: DINT;
		SubCmd 	: DINT;
		ParaValue 	: DINT;
	END_VAR
	VAR_OUTPUT
		Retcode 	: DINT;
	END_VAR
VAR
	pConn       : ^_CONNECTION;
END_VAR

  Retcode := TCP_SVR_NO_ERROR;

  if (CheckSocketValid(dSock, (#pConn)$^pVoid) = true) then
    if (pConn <> NIL) then
      case Cmd of
        (*================================================================*)
        SVR_TCP_CMD_SETSOCKOPT:
        (*================================================================*)
          case SubCmd of
            (*==================================================*)
            SVR_TCP_SOCKOPT_NAGLE:
            (*==================================================*)
              if (ParaValue = 0) then
                if (pConn^.ConnSockOpt.Nagle = true) then
                  AP_SemaWait(AP_SemaSockOpt);
                  pConn^.ConnSockOpt.Nagle := false;
                  pConn^.bdSettings.SockOptChanged := true;
                  AP_SemaSignal(AP_SemaSockOpt);
                end_if;
              else
                if (pConn^.ConnSockOpt.Nagle = false) then
                  AP_SemaWait(AP_SemaSockOpt);
                  pConn^.ConnSockOpt.Nagle := true;
                  pConn^.bdSettings.SockOptChanged := true;
                  AP_SemaSignal(AP_SemaSockOpt);
                end_if;
              end_if;
            (*==================================================*)
            SVR_TCP_SOCKOPT_KEEPALIVE:
            (*==================================================*)
              if (ParaValue = 0) then
                if (pConn^.ConnSockOpt.KeepAlive = true) then
                  AP_SemaWait(AP_SemaSockOpt);
                  pConn^.ConnSockOpt.KeepAlive := false;
                  pConn^.bdSettings.SockOptChanged := true;
                  AP_SemaSignal(AP_SemaSockOpt);
                end_if;
              else
                if (pConn^.ConnSockOpt.KeepAlive = false) then
                  AP_SemaWait(AP_SemaSockOpt);
                  pConn^.ConnSockOpt.KeepAlive := true;
                  pConn^.bdSettings.SockOptChanged := true;
                  AP_SemaSignal(AP_SemaSockOpt);
                end_if;
              end_if;
            (*==================================================*)
            SVR_TCP_SOCKOPT_DELAYEDACK:
            (*==================================================*)
              if (ParaValue = 0) then
                if (pConn^.ConnSockOpt.DelayedAck = true) then
                  AP_SemaWait(AP_SemaSockOpt);
                  pConn^.ConnSockOpt.DelayedAck := false;
                  pConn^.bdSettings.SockOptChanged := true;
                  AP_SemaSignal(AP_SemaSockOpt);
                end_if;
              else
                if (pConn^.ConnSockOpt.DelayedAck = false) then
                  AP_SemaWait(AP_SemaSockOpt);
                  pConn^.ConnSockOpt.DelayedAck := true;
                  pConn^.bdSettings.SockOptChanged := true;
                  AP_SemaSignal(AP_SemaSockOpt);
                end_if;
              end_if;
            (*==================================================*)
            SVR_TCP_SOCKOPT_REUSEADDR:
            (*==================================================*)
              if (ParaValue = 0) then
                if (pConn^.ConnSockOpt.ReuseAddr = true) then
                  AP_SemaWait(AP_SemaSockOpt);
                  pConn^.ConnSockOpt.ReuseAddr := false;
                  pConn^.bdSettings.SockOptChanged := true;
                  AP_SemaSignal(AP_SemaSockOpt);
                end_if;
              else
                if (pConn^.ConnSockOpt.ReuseAddr = false) then
                  AP_SemaWait(AP_SemaSockOpt);
                  pConn^.ConnSockOpt.ReuseAddr := true;
                  pConn^.bdSettings.SockOptChanged := true;
                  AP_SemaSignal(AP_SemaSockOpt);
                end_if;
              end_if;
            (*==================================================*)
            else // - INVALID SUB COMMAND
            (*==================================================*)
              Retcode := TCP_SVR_ERR_SET_PARA_INVALID_SUB_CMD;
          end_case;

        (*================================================================*)
        SVR_TCP_CMD_KEEPALIVEPARA: // - ASYNC TASK PRIORITY
        (*================================================================*)
          case SubCmd of
            (*==================================================*)
            SVR_TCP_KEEPALIVE_KEEPIDLE:
            (*==================================================*)
              AP_SemaWait(AP_SemaSockOpt);
              pConn^.KeepAlivePara.keepIDLE    := ParaValue;
              pConn^.bdSettings.SockOptChanged := true;
              AP_SemaSignal(AP_SemaSockOpt);
            (*==================================================*)
            SVR_TCP_KEEPALIVE_KEEPINTVL:
            (*==================================================*)
              AP_SemaWait(AP_SemaSockOpt);
              pConn^.KeepAlivePara.keepINTVL   := ParaValue;
              pConn^.bdSettings.SockOptChanged := true;
              AP_SemaSignal(AP_SemaSockOpt);
            (*==================================================*)
            SVR_TCP_KEEPALIVE_KEEPCNT:
            (*==================================================*)
              AP_SemaWait(AP_SemaSockOpt);
              pConn^.KeepAlivePara.keepCNT     := ParaValue;
              pConn^.bdSettings.SockOptChanged := true;
              AP_SemaSignal(AP_SemaSockOpt);
            (*==================================================*)
            else // - INVALID SUB COMMAND
            (*==================================================*)
              Retcode := TCP_SVR_ERR_SET_PARA_INVALID_SUB_CMD;
          end_case;
